ACTION act_Oper:
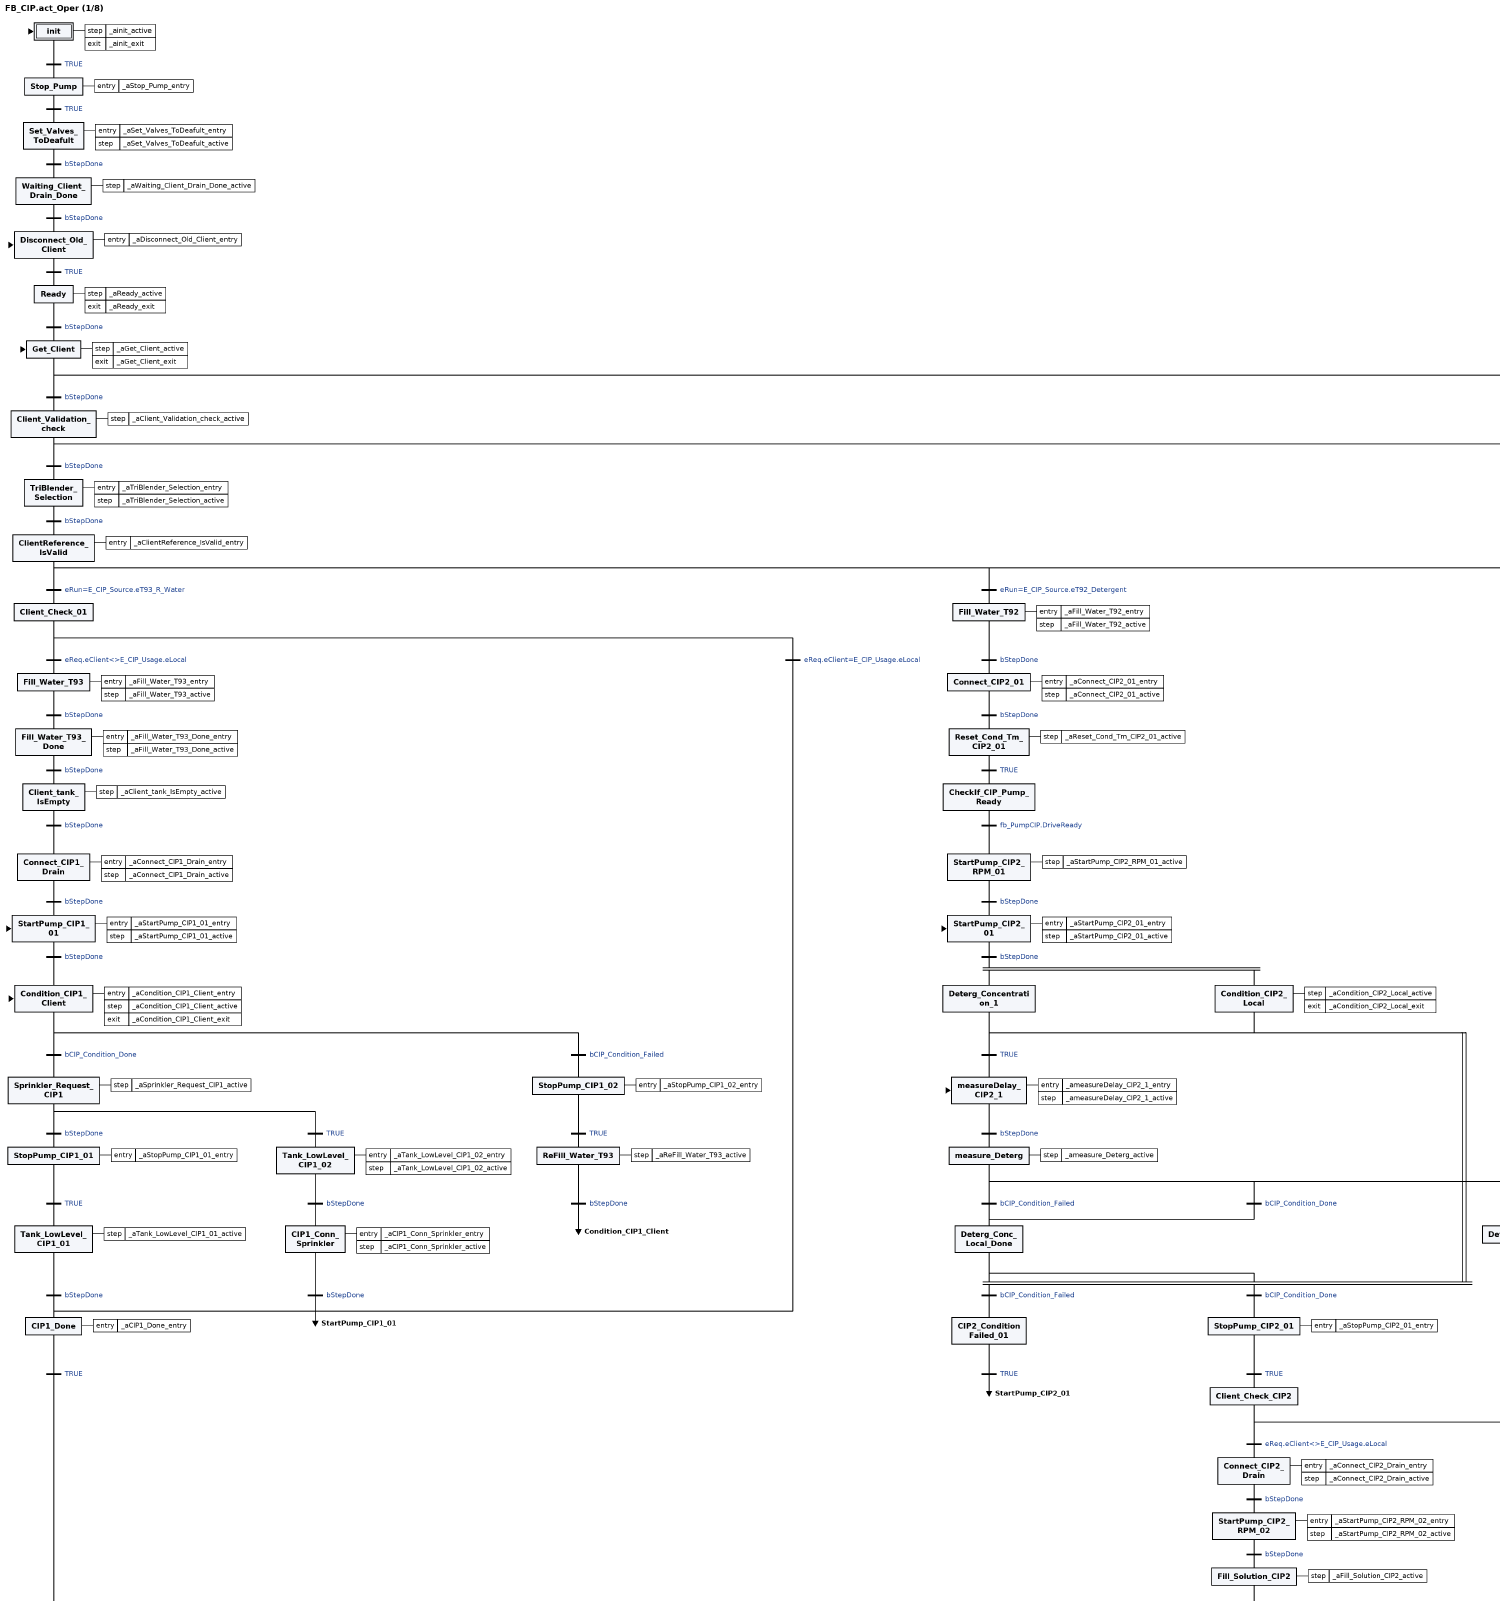
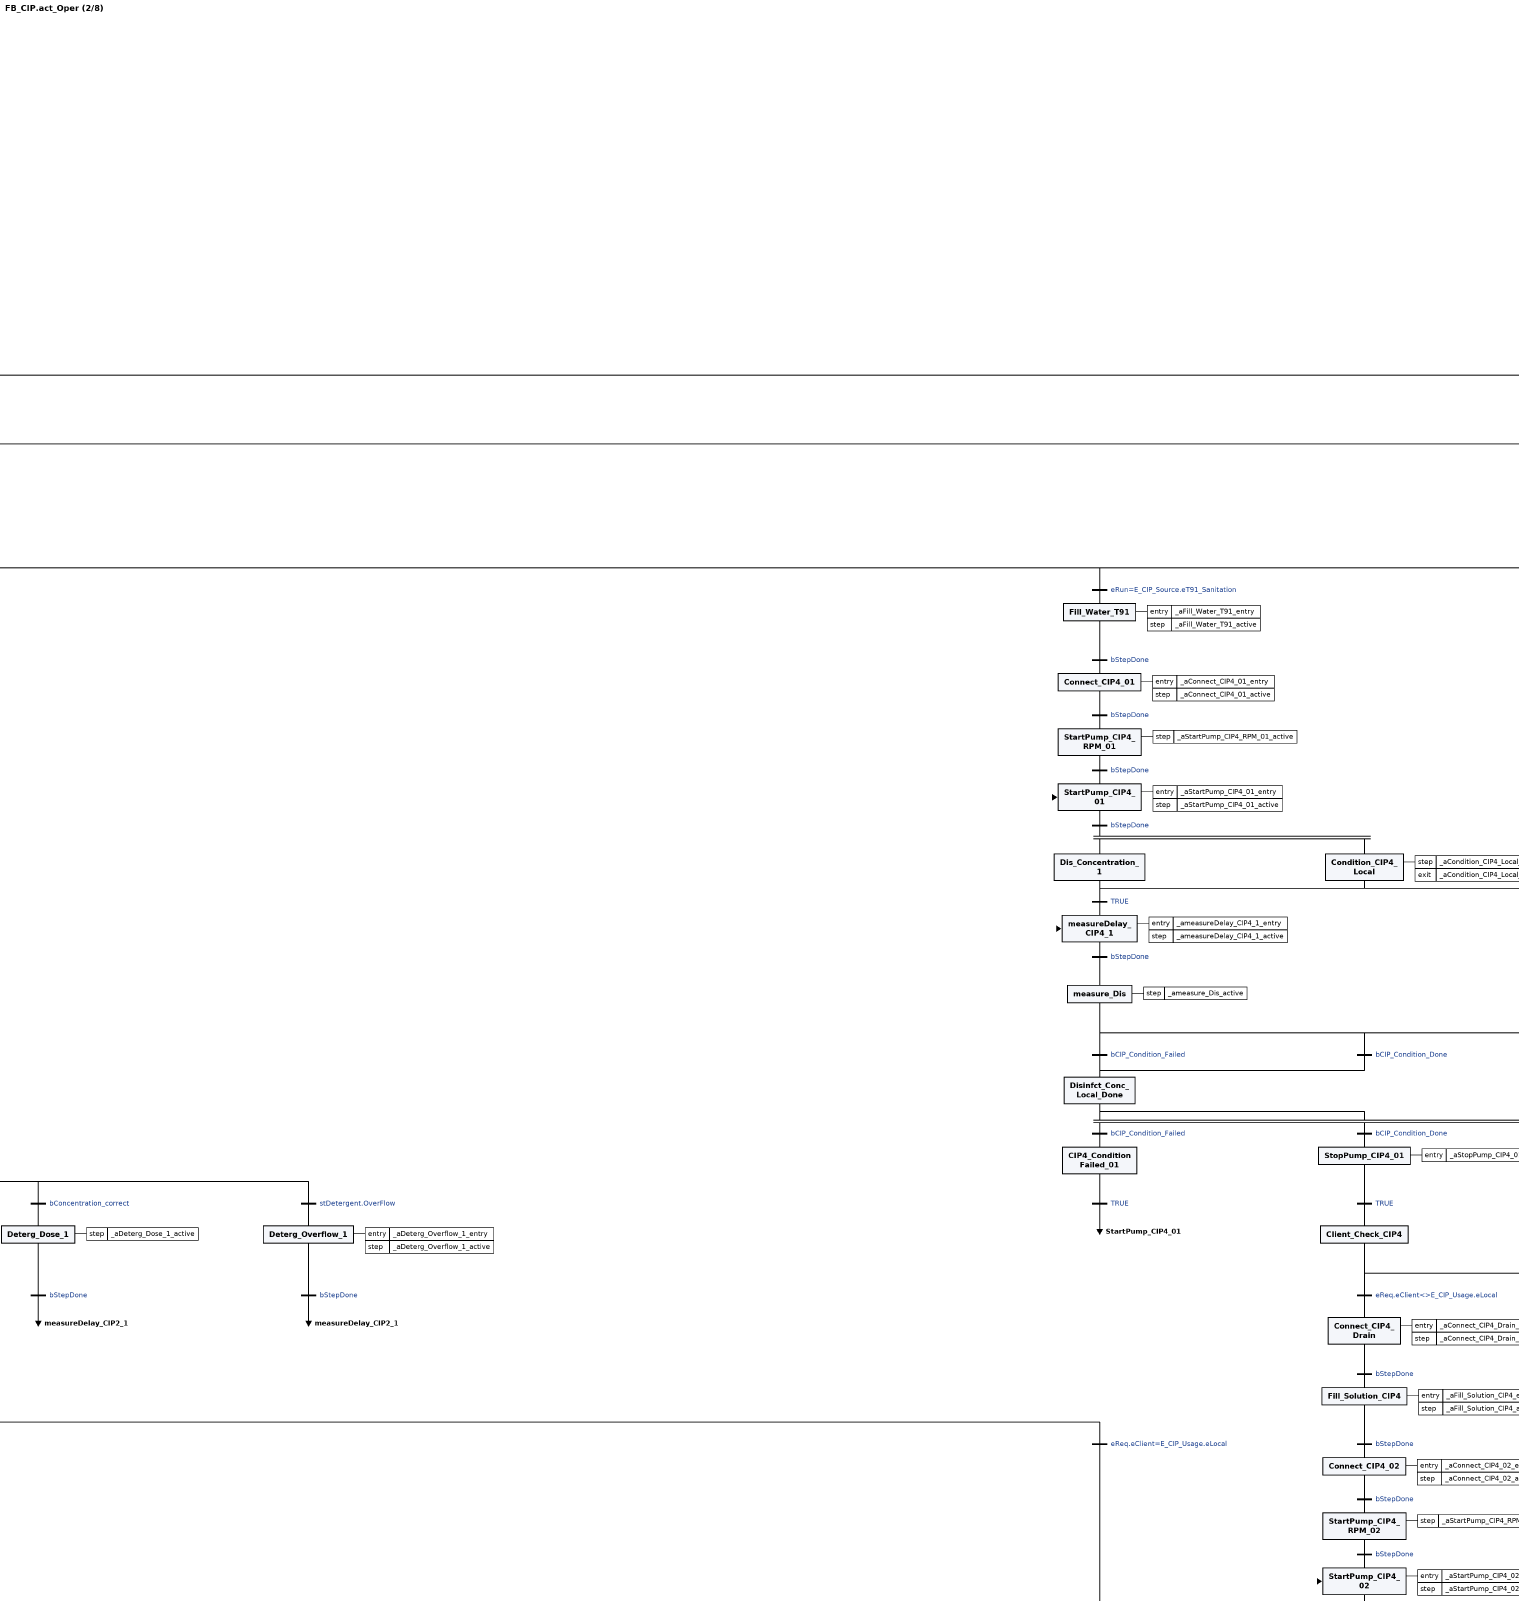
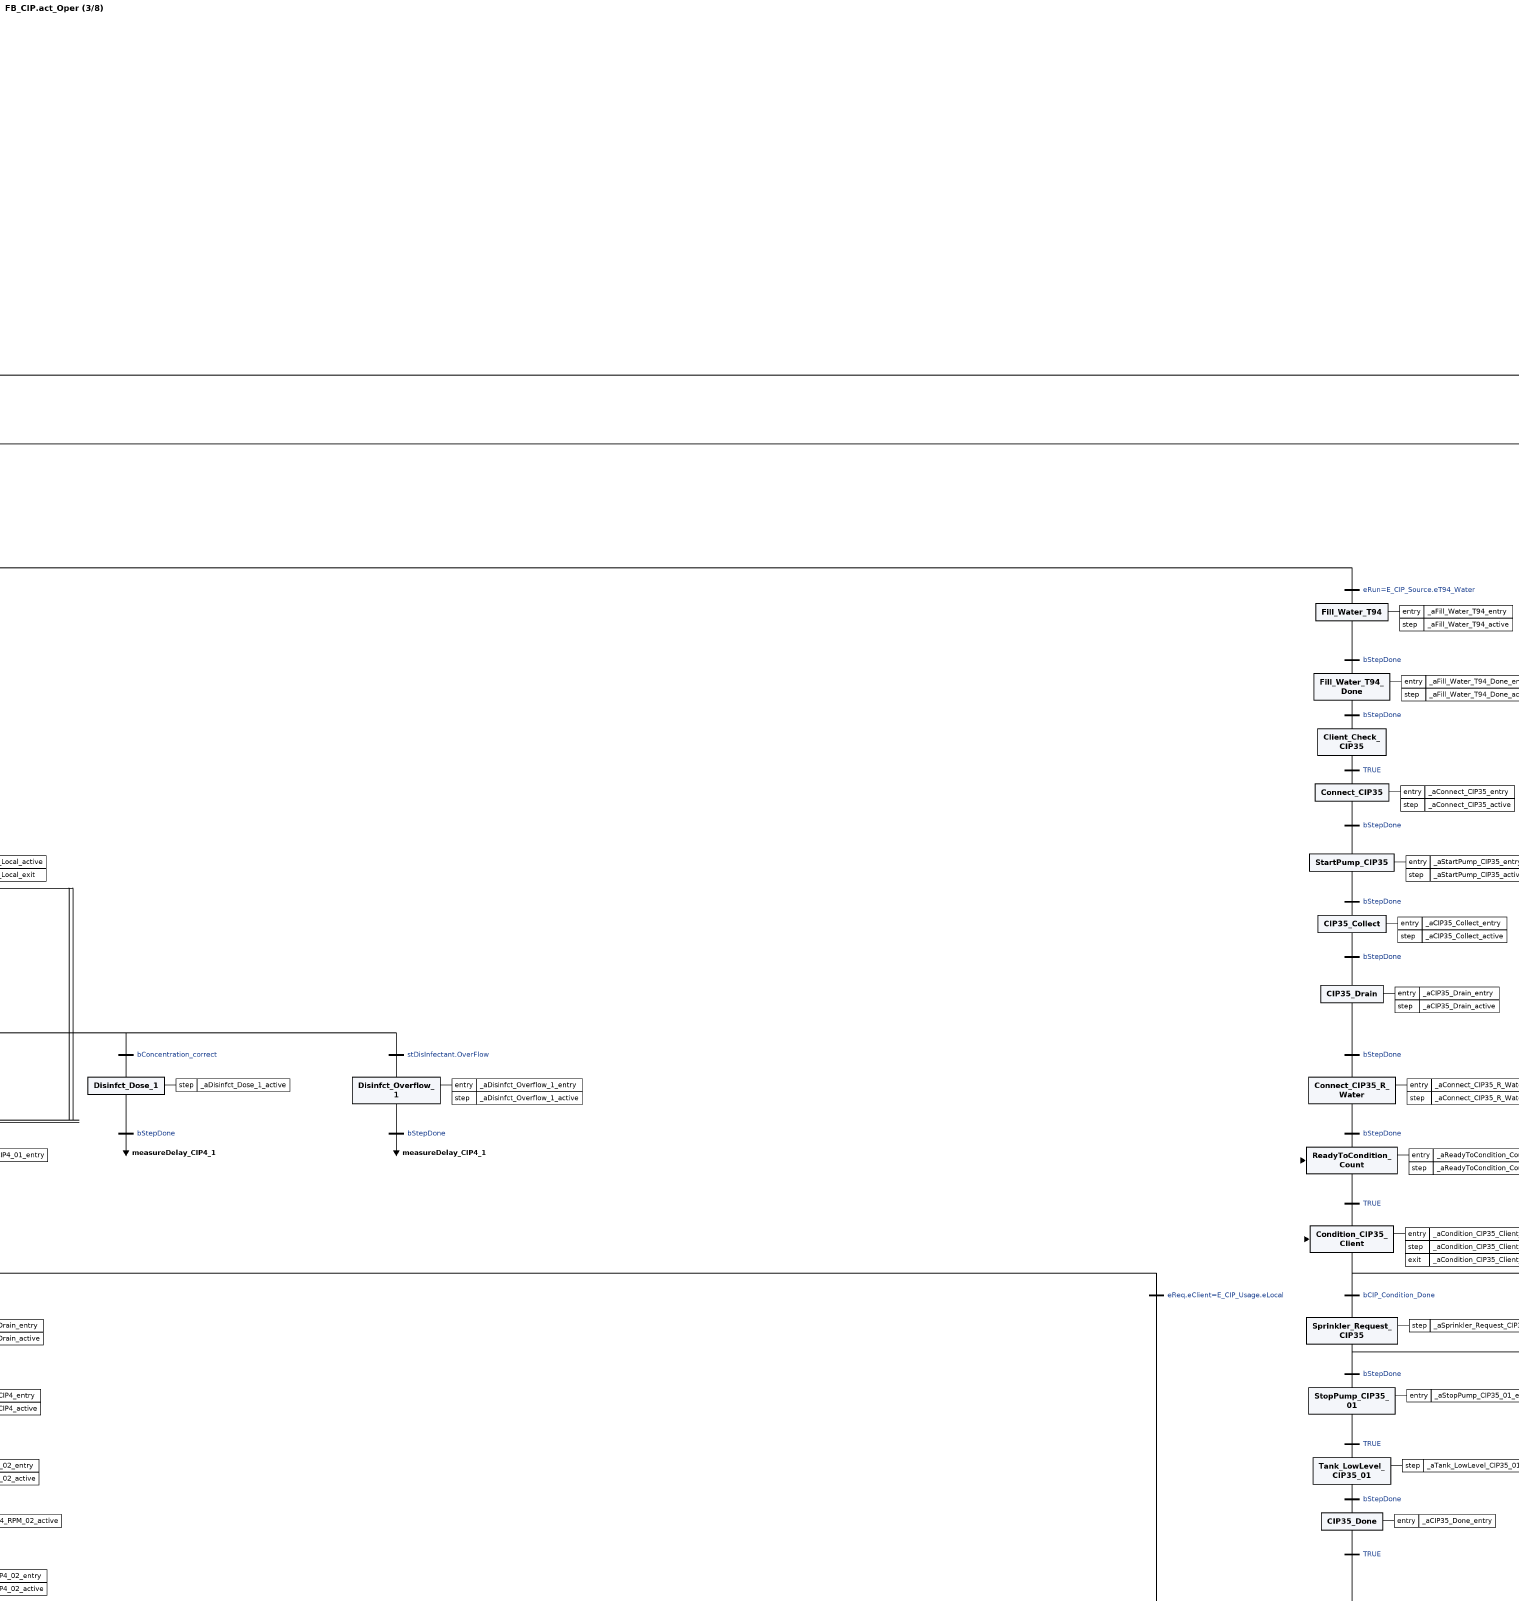
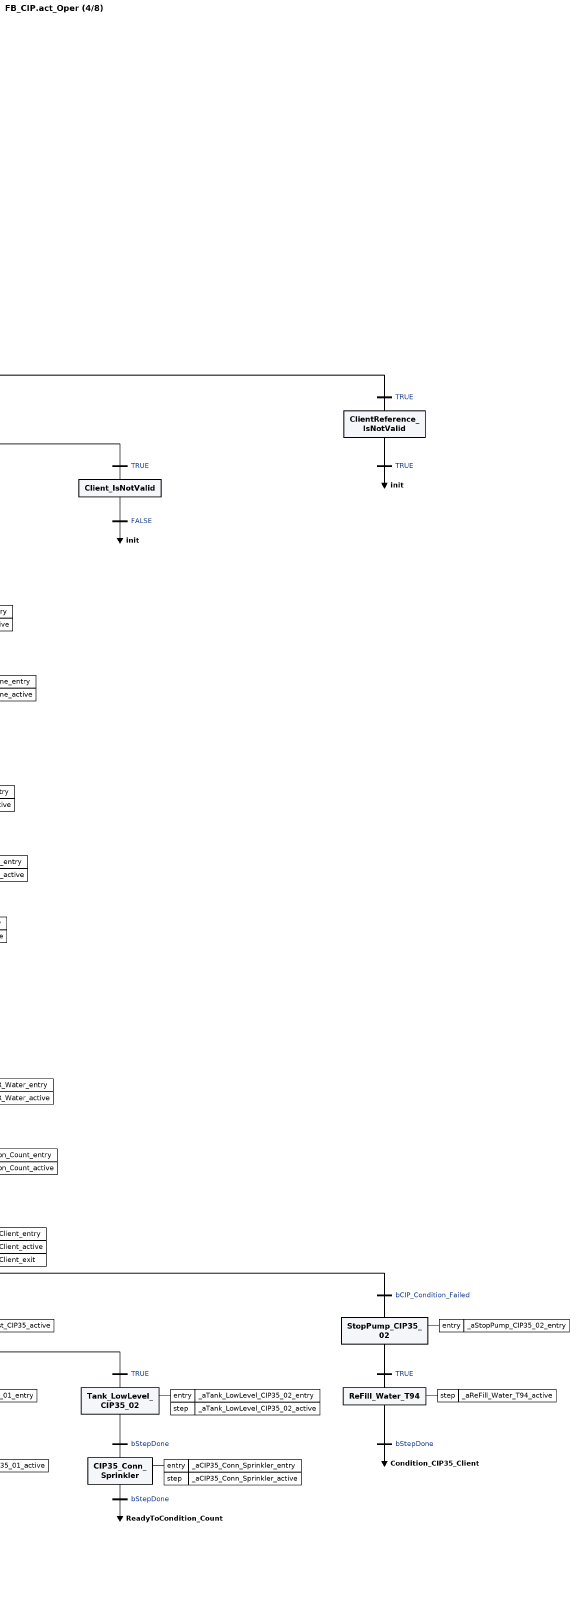
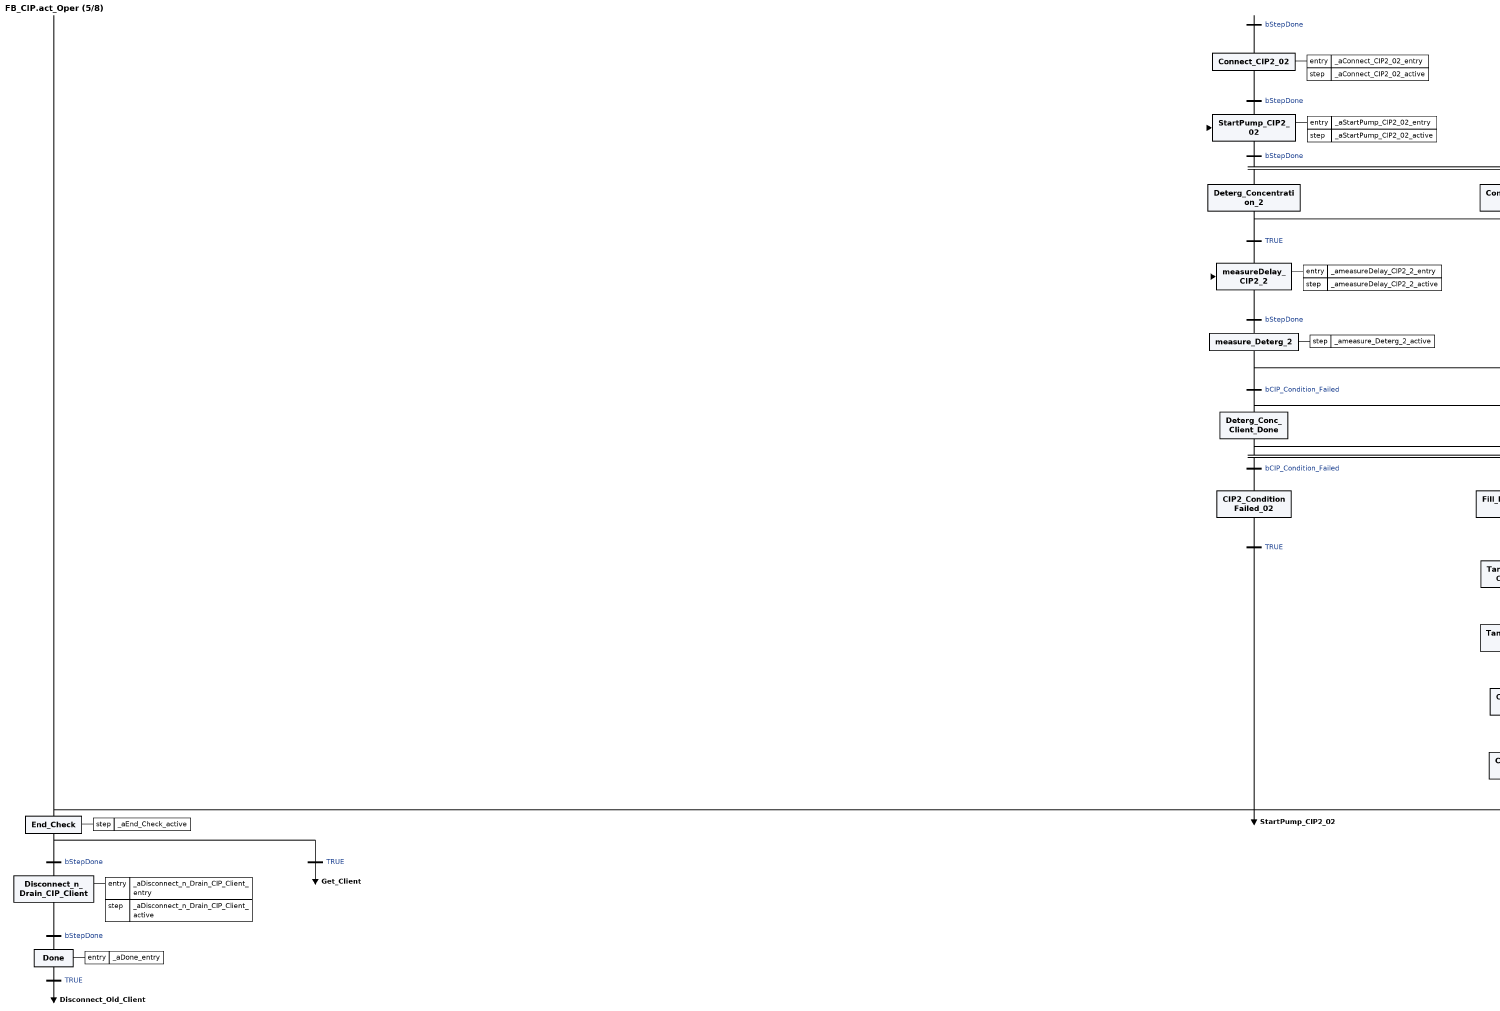
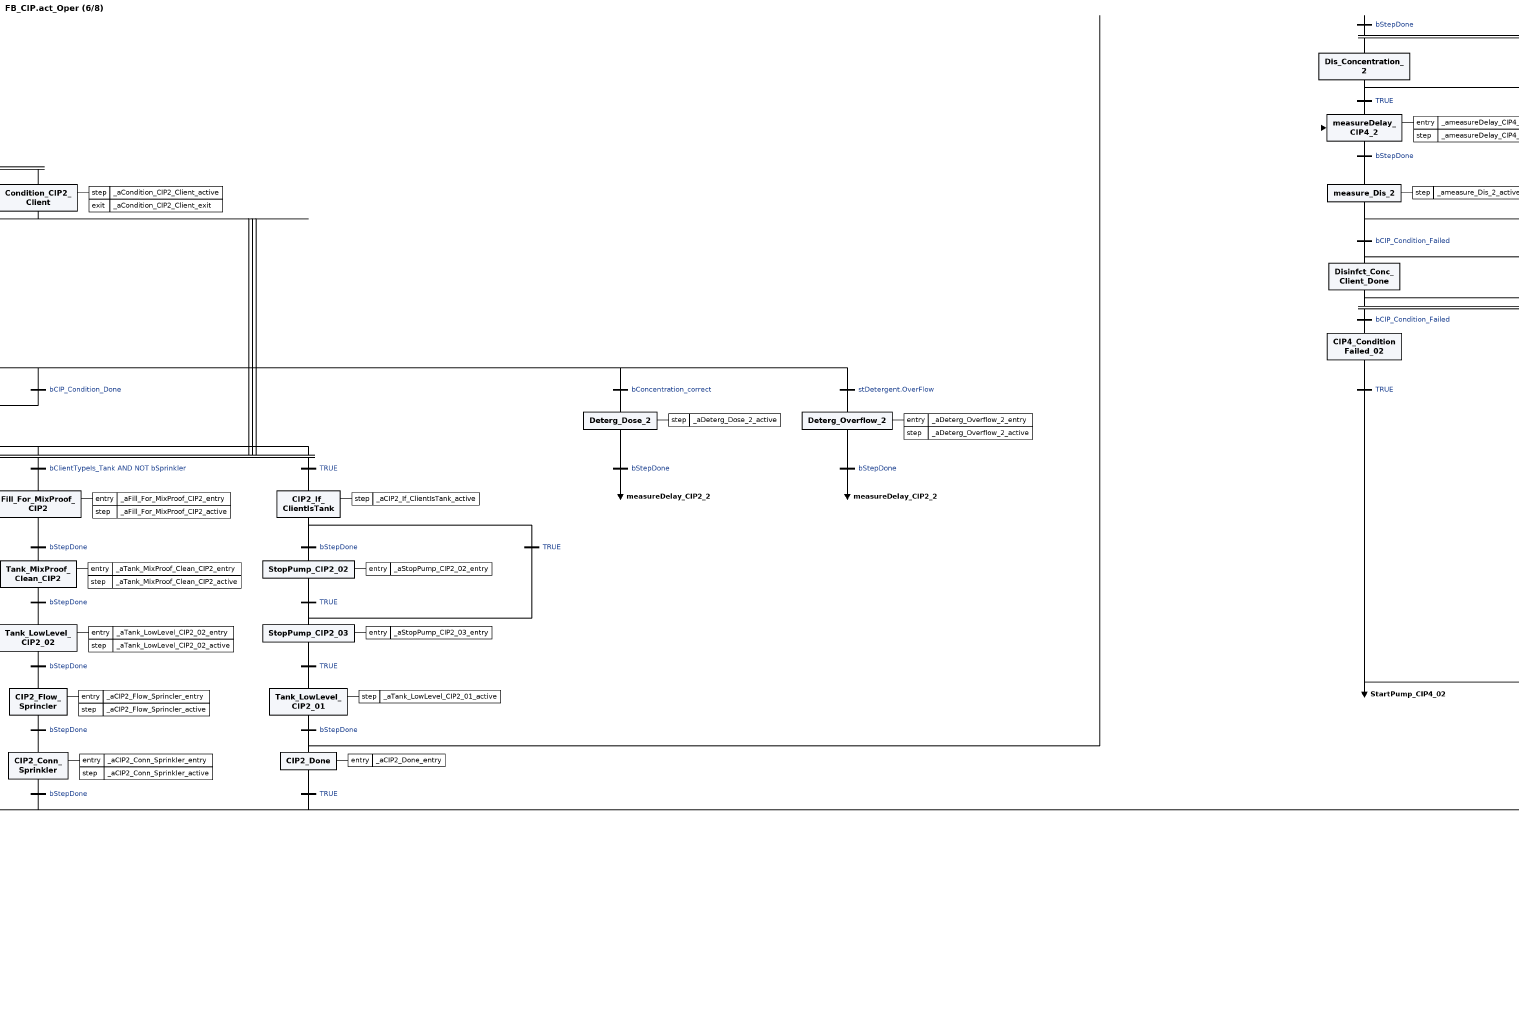
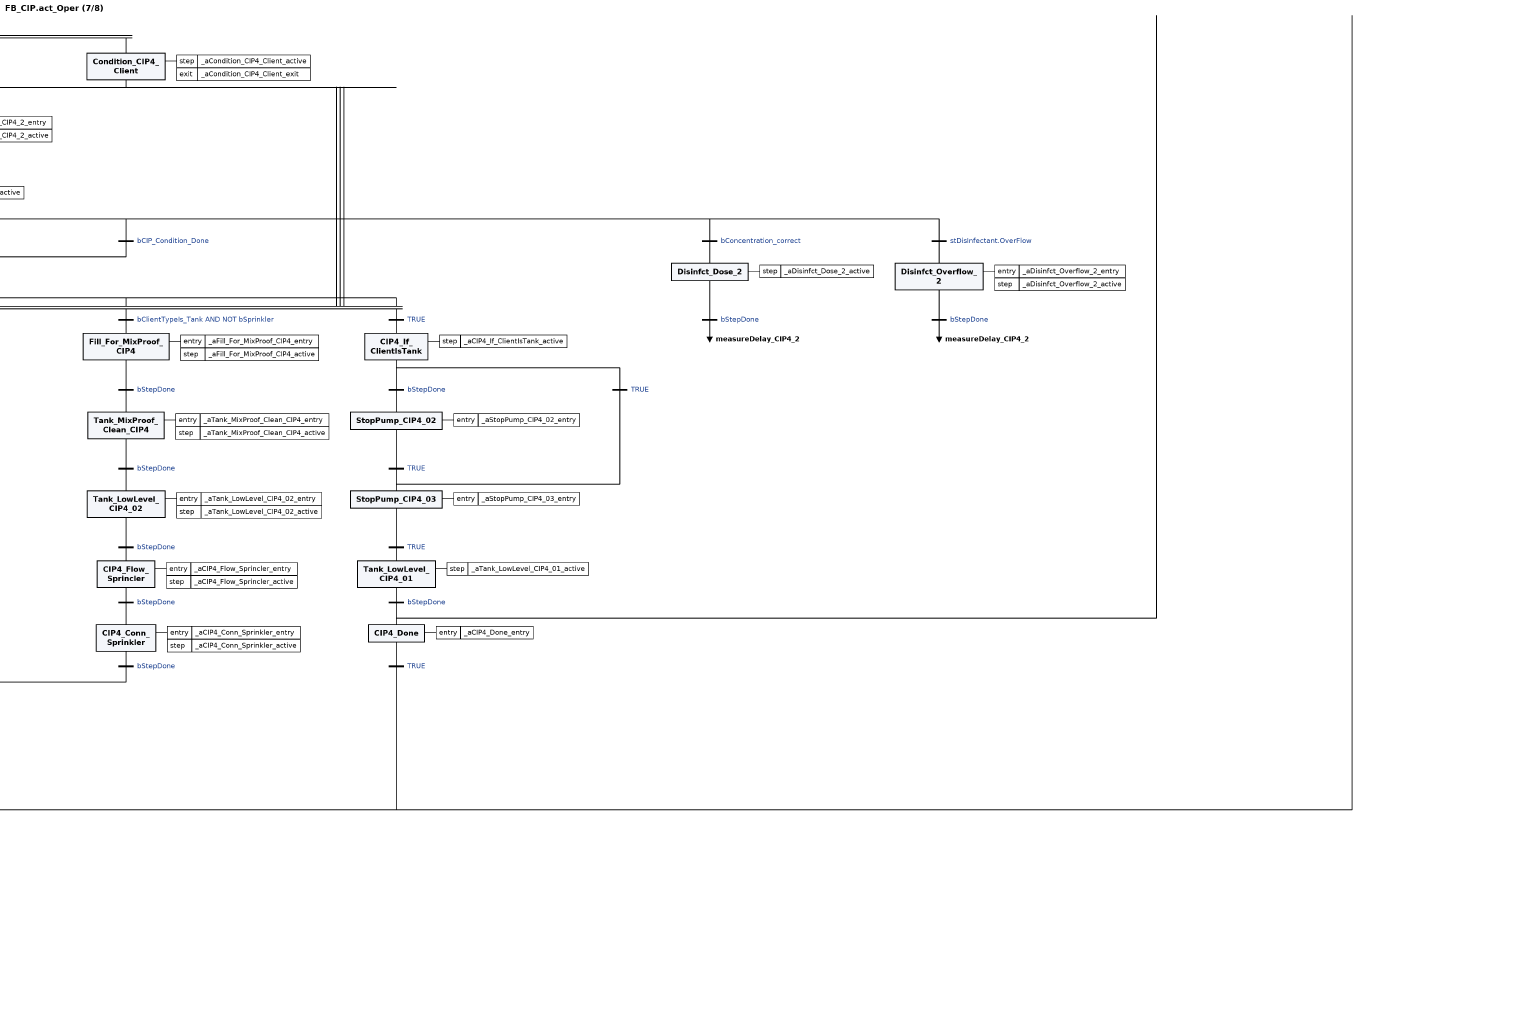
INITIAL_STEP init:
    _ainit_active(N);  // step action
    _ainit_exit(P0);  // exit action
END_STEP
TRANSITION FROM init TO Stop_Pump
    := TRUE;
END_TRANSITION
STEP Stop_Pump:
    _aStop_Pump_entry(P1);  // entry action
END_STEP
TRANSITION FROM Stop_Pump TO Set_Valves_ToDeafult
    := TRUE;
END_TRANSITION
STEP Set_Valves_ToDeafult:  // min time T#0.1s
    _aSet_Valves_ToDeafult_entry(P1);  // entry action
    _aSet_Valves_ToDeafult_active(N);  // step action
END_STEP
TRANSITION FROM Set_Valves_ToDeafult TO Waiting_Client_Drain_Done
    := bStepDone;
END_TRANSITION
STEP Waiting_Client_Drain_Done:  // min time T#0.1s
    _aWaiting_Client_Drain_Done_active(N);  // step action
END_STEP
TRANSITION FROM Waiting_Client_Drain_Done TO Disconnect_Old_Client
    := bStepDone;
END_TRANSITION
STEP Disconnect_Old_Client:
    _aDisconnect_Old_Client_entry(P1);  // entry action
END_STEP
TRANSITION FROM Disconnect_Old_Client TO Ready
    := TRUE;
END_TRANSITION
STEP Ready:
    _aReady_active(N);  // step action
    _aReady_exit(P0);  // exit action
END_STEP
TRANSITION FROM Ready TO Get_Client
    := bStepDone;
END_TRANSITION
STEP Get_Client:  // max time T#0.1s
    _aGet_Client_active(N);  // step action
    _aGet_Client_exit(P0);  // exit action
END_STEP
TRANSITION FROM Get_Client TO Client_Validation_check
    := bStepDone;
END_TRANSITION
TRANSITION FROM Get_Client TO ClientReference_IsNotValid
    := TRUE;
END_TRANSITION
STEP ClientReference_IsNotValid:  // min time T#2s
END_STEP
TRANSITION FROM ClientReference_IsNotValid TO init
    := TRUE;
END_TRANSITION
STEP Client_Validation_check:
    _aClient_Validation_check_active(N);  // step action
END_STEP
TRANSITION FROM Client_Validation_check TO TriBlender_Selection
    := bStepDone;
END_TRANSITION
STEP TriBlender_Selection:
    _aTriBlender_Selection_entry(P1);  // entry action
    _aTriBlender_Selection_active(N);  // step action
END_STEP
TRANSITION FROM TriBlender_Selection TO ClientReference_IsValid
    := bStepDone;
END_TRANSITION
TRANSITION FROM Client_Validation_check TO Client_IsNotValid
    := TRUE;
END_TRANSITION
STEP Client_IsNotValid:  // min time T#2s
END_STEP
TRANSITION FROM Client_IsNotValid TO init
    := FALSE;
END_TRANSITION
STEP ClientReference_IsValid:
    _aClientReference_IsValid_entry(P1);  // entry action
END_STEP
TRANSITION FROM ClientReference_IsValid TO Client_Check_01
    := eRun=E_CIP_Source.eT93_R_Water;
END_TRANSITION
// macro R_Water begins
STEP Client_Check_01:
END_STEP
TRANSITION FROM Client_Check_01 TO Fill_Water_T93
    := eReq.eClient<>E_CIP_Usage.eLocal;
END_TRANSITION
STEP Fill_Water_T93:
    _aFill_Water_T93_entry(P1);  // entry action
    _aFill_Water_T93_active(N);  // step action
END_STEP
TRANSITION FROM Fill_Water_T93 TO Fill_Water_T93_Done
    := bStepDone;
END_TRANSITION
STEP Fill_Water_T93_Done:
    _aFill_Water_T93_Done_entry(P1);  // entry action
    _aFill_Water_T93_Done_active(N);  // step action
END_STEP
TRANSITION FROM Fill_Water_T93_Done TO Client_tank_IsEmpty
    := bStepDone;
END_TRANSITION
STEP Client_tank_IsEmpty:  // min time T#5s
    _aClient_tank_IsEmpty_active(N);  // step action
END_STEP
TRANSITION FROM Client_tank_IsEmpty TO Connect_CIP1_Drain
    := bStepDone;
END_TRANSITION
STEP Connect_CIP1_Drain:
    _aConnect_CIP1_Drain_entry(P1);  // entry action
    _aConnect_CIP1_Drain_active(N);  // step action
END_STEP
TRANSITION FROM Connect_CIP1_Drain TO StartPump_CIP1_01
    := bStepDone;
END_TRANSITION
STEP StartPump_CIP1_01:
    _aStartPump_CIP1_01_entry(P1);  // entry action
    _aStartPump_CIP1_01_active(N);  // step action
END_STEP
TRANSITION FROM StartPump_CIP1_01 TO Condition_CIP1_Client
    := bStepDone;
END_TRANSITION
STEP Condition_CIP1_Client:
    _aCondition_CIP1_Client_entry(P1);  // entry action
    _aCondition_CIP1_Client_active(N);  // step action
    _aCondition_CIP1_Client_exit(P0);  // exit action
END_STEP
TRANSITION FROM Condition_CIP1_Client TO Sprinkler_Request_CIP1
    := bCIP_Condition_Done;
END_TRANSITION
STEP Sprinkler_Request_CIP1:
    _aSprinkler_Request_CIP1_active(N);  // step action
END_STEP
TRANSITION FROM Sprinkler_Request_CIP1 TO StopPump_CIP1_01
    := bStepDone;
END_TRANSITION
STEP StopPump_CIP1_01:
    _aStopPump_CIP1_01_entry(P1);  // entry action
END_STEP
TRANSITION FROM StopPump_CIP1_01 TO Tank_LowLevel_CIP1_01
    := TRUE;
END_TRANSITION
STEP Tank_LowLevel_CIP1_01:
    _aTank_LowLevel_CIP1_01_active(N);  // step action
END_STEP
TRANSITION FROM Tank_LowLevel_CIP1_01 TO CIP1_Done
    := bStepDone;
END_TRANSITION
TRANSITION FROM Sprinkler_Request_CIP1 TO Tank_LowLevel_CIP1_02
    := TRUE;
END_TRANSITION
STEP Tank_LowLevel_CIP1_02:
    _aTank_LowLevel_CIP1_02_entry(P1);  // entry action
    _aTank_LowLevel_CIP1_02_active(N);  // step action
END_STEP
TRANSITION FROM Tank_LowLevel_CIP1_02 TO CIP1_Conn_Sprinkler
    := bStepDone;
END_TRANSITION
STEP CIP1_Conn_Sprinkler:
    _aCIP1_Conn_Sprinkler_entry(P1);  // entry action
    _aCIP1_Conn_Sprinkler_active(N);  // step action
END_STEP
TRANSITION FROM CIP1_Conn_Sprinkler TO StartPump_CIP1_01
    := bStepDone;
END_TRANSITION
TRANSITION FROM Condition_CIP1_Client TO StopPump_CIP1_02
    := bCIP_Condition_Failed;
END_TRANSITION
STEP StopPump_CIP1_02:
    _aStopPump_CIP1_02_entry(P1);  // entry action
END_STEP
TRANSITION FROM StopPump_CIP1_02 TO ReFill_Water_T93
    := TRUE;
END_TRANSITION
STEP ReFill_Water_T93:
    _aReFill_Water_T93_active(N);  // step action
END_STEP
TRANSITION FROM ReFill_Water_T93 TO Condition_CIP1_Client
    := bStepDone;
END_TRANSITION
TRANSITION FROM Client_Check_01 TO CIP1_Done
    := eReq.eClient=E_CIP_Usage.eLocal;
END_TRANSITION
STEP CIP1_Done:  // min time T#2s
    _aCIP1_Done_entry(P1);  // entry action
END_STEP
TRANSITION FROM CIP1_Done TO End_Check
    := TRUE;
END_TRANSITION
TRANSITION FROM ClientReference_IsValid TO Fill_Water_T92
    := eRun=E_CIP_Source.eT92_Detergent;
END_TRANSITION
// macro Detergent begins
STEP Fill_Water_T92:
    _aFill_Water_T92_entry(P1);  // entry action
    _aFill_Water_T92_active(N);  // step action
END_STEP
TRANSITION FROM Fill_Water_T92 TO Connect_CIP2_01
    := bStepDone;
END_TRANSITION
STEP Connect_CIP2_01:
    _aConnect_CIP2_01_entry(P1);  // entry action
    _aConnect_CIP2_01_active(N);  // step action
END_STEP
TRANSITION FROM Connect_CIP2_01 TO Reset_Cond_Tm_CIP2_01
    := bStepDone;
END_TRANSITION
STEP Reset_Cond_Tm_CIP2_01:
    _aReset_Cond_Tm_CIP2_01_active(N);  // step action
END_STEP
TRANSITION FROM Reset_Cond_Tm_CIP2_01 TO CheckIf_CIP_Pump_Ready
    := TRUE;
END_TRANSITION
STEP CheckIf_CIP_Pump_Ready:
END_STEP
TRANSITION FROM CheckIf_CIP_Pump_Ready TO StartPump_CIP2_RPM_01
    := fb_PumpCIP.DriveReady;
END_TRANSITION
STEP StartPump_CIP2_RPM_01:
    _aStartPump_CIP2_RPM_01_active(N);  // step action
END_STEP
TRANSITION FROM StartPump_CIP2_RPM_01 TO StartPump_CIP2_01
    := bStepDone;
END_TRANSITION
STEP StartPump_CIP2_01:  // min time T#2s
    _aStartPump_CIP2_01_entry(P1);  // entry action
    _aStartPump_CIP2_01_active(N);  // step action
END_STEP
TRANSITION FROM StartPump_CIP2_01 TO (Deterg_Concentration_1, Condition_CIP2_Local)
    := bStepDone;
END_TRANSITION
STEP Deterg_Concentration_1:
END_STEP
TRANSITION FROM Deterg_Concentration_1 TO measureDelay_CIP2_1
    := TRUE;
END_TRANSITION
STEP measureDelay_CIP2_1:
    _ameasureDelay_CIP2_1_entry(P1);  // entry action
    _ameasureDelay_CIP2_1_active(N);  // step action
END_STEP
TRANSITION FROM measureDelay_CIP2_1 TO measure_Deterg
    := bStepDone;
END_TRANSITION
STEP measure_Deterg:  // min time t#1s
    _ameasure_Deterg_active(N);  // step action
END_STEP
TRANSITION FROM measure_Deterg TO Deterg_Conc_Local_Done
    := bCIP_Condition_Failed;
END_TRANSITION
TRANSITION FROM measure_Deterg TO Deterg_Conc_Local_Done
    := bCIP_Condition_Done;
END_TRANSITION
TRANSITION FROM measure_Deterg TO Deterg_Dose_1
    := bConcentration_correct;
END_TRANSITION
STEP Deterg_Dose_1:
    _aDeterg_Dose_1_active(N);  // step action
END_STEP
TRANSITION FROM Deterg_Dose_1 TO measureDelay_CIP2_1
    := bStepDone;
END_TRANSITION
TRANSITION FROM measure_Deterg TO Deterg_Overflow_1
    := stDetergent.OverFlow;
END_TRANSITION
STEP Deterg_Overflow_1:
    _aDeterg_Overflow_1_entry(P1);  // entry action
    _aDeterg_Overflow_1_active(N);  // step action
END_STEP
TRANSITION FROM Deterg_Overflow_1 TO measureDelay_CIP2_1
    := bStepDone;
END_TRANSITION
STEP Deterg_Conc_Local_Done:
END_STEP
STEP Condition_CIP2_Local:
    _aCondition_CIP2_Local_active(N);  // step action
    _aCondition_CIP2_Local_exit(P0);  // exit action
END_STEP
TRANSITION FROM (Deterg_Conc_Local_Done, Condition_CIP2_Local) TO CIP2_ConditionFailed_01
    := bCIP_Condition_Failed;
END_TRANSITION
STEP CIP2_ConditionFailed_01:
END_STEP
TRANSITION FROM CIP2_ConditionFailed_01 TO StartPump_CIP2_01
    := TRUE;
END_TRANSITION
TRANSITION FROM (Deterg_Conc_Local_Done, Condition_CIP2_Local) TO StopPump_CIP2_01
    := bCIP_Condition_Done;
END_TRANSITION
STEP StopPump_CIP2_01:
    _aStopPump_CIP2_01_entry(P1);  // entry action
END_STEP
TRANSITION FROM StopPump_CIP2_01 TO Client_Check_CIP2
    := TRUE;
END_TRANSITION
STEP Client_Check_CIP2:
END_STEP
TRANSITION FROM Client_Check_CIP2 TO Connect_CIP2_Drain
    := eReq.eClient<>E_CIP_Usage.eLocal;
END_TRANSITION
STEP Connect_CIP2_Drain:
    _aConnect_CIP2_Drain_entry(P1);  // entry action
    _aConnect_CIP2_Drain_active(N);  // step action
END_STEP
TRANSITION FROM Connect_CIP2_Drain TO StartPump_CIP2_RPM_02
    := bStepDone;
END_TRANSITION
STEP StartPump_CIP2_RPM_02:
    _aStartPump_CIP2_RPM_02_entry(P1);  // entry action
    _aStartPump_CIP2_RPM_02_active(N);  // step action
END_STEP
TRANSITION FROM StartPump_CIP2_RPM_02 TO Fill_Solution_CIP2
    := bStepDone;
END_TRANSITION
STEP Fill_Solution_CIP2:
    _aFill_Solution_CIP2_active(N);  // step action
END_STEP
TRANSITION FROM Fill_Solution_CIP2 TO Connect_CIP2_02
    := bStepDone;
END_TRANSITION
STEP Connect_CIP2_02:
    _aConnect_CIP2_02_entry(P1);  // entry action
    _aConnect_CIP2_02_active(N);  // step action
END_STEP
TRANSITION FROM Connect_CIP2_02 TO StartPump_CIP2_02
    := bStepDone;
END_TRANSITION
STEP StartPump_CIP2_02:  // min time T#2s
    _aStartPump_CIP2_02_entry(P1);  // entry action
    _aStartPump_CIP2_02_active(N);  // step action
END_STEP
TRANSITION FROM StartPump_CIP2_02 TO (Deterg_Concentration_2, Condition_CIP2_Client)
    := bStepDone;
END_TRANSITION
STEP Deterg_Concentration_2:
END_STEP
TRANSITION FROM Deterg_Concentration_2 TO measureDelay_CIP2_2
    := TRUE;
END_TRANSITION
STEP measureDelay_CIP2_2:
    _ameasureDelay_CIP2_2_entry(P1);  // entry action
    _ameasureDelay_CIP2_2_active(N);  // step action
END_STEP
TRANSITION FROM measureDelay_CIP2_2 TO measure_Deterg_2
    := bStepDone;
END_TRANSITION
STEP measure_Deterg_2:  // min time t#1s
    _ameasure_Deterg_2_active(N);  // step action
END_STEP
TRANSITION FROM measure_Deterg_2 TO Deterg_Conc_Client_Done
    := bCIP_Condition_Failed;
END_TRANSITION
TRANSITION FROM measure_Deterg_2 TO Deterg_Conc_Client_Done
    := bCIP_Condition_Done;
END_TRANSITION
TRANSITION FROM measure_Deterg_2 TO Deterg_Dose_2
    := bConcentration_correct;
END_TRANSITION
STEP Deterg_Dose_2:
    _aDeterg_Dose_2_active(N);  // step action
END_STEP
TRANSITION FROM Deterg_Dose_2 TO measureDelay_CIP2_2
    := bStepDone;
END_TRANSITION
TRANSITION FROM measure_Deterg_2 TO Deterg_Overflow_2
    := stDetergent.OverFlow;
END_TRANSITION
STEP Deterg_Overflow_2:
    _aDeterg_Overflow_2_entry(P1);  // entry action
    _aDeterg_Overflow_2_active(N);  // step action
END_STEP
TRANSITION FROM Deterg_Overflow_2 TO measureDelay_CIP2_2
    := bStepDone;
END_TRANSITION
STEP Deterg_Conc_Client_Done:
END_STEP
STEP Condition_CIP2_Client:
    _aCondition_CIP2_Client_active(N);  // step action
    _aCondition_CIP2_Client_exit(P0);  // exit action
END_STEP
TRANSITION FROM (Deterg_Conc_Client_Done, Condition_CIP2_Client) TO CIP2_ConditionFailed_02
    := bCIP_Condition_Failed;
END_TRANSITION
STEP CIP2_ConditionFailed_02:
END_STEP
TRANSITION FROM CIP2_ConditionFailed_02 TO StartPump_CIP2_02
    := TRUE;
END_TRANSITION
TRANSITION FROM (Deterg_Conc_Client_Done, Condition_CIP2_Client) TO Fill_For_MixProof_CIP2
    := bClientTypeIs_Tank AND NOT bSprinkler;
END_TRANSITION
STEP Fill_For_MixProof_CIP2:
    _aFill_For_MixProof_CIP2_entry(P1);  // entry action
    _aFill_For_MixProof_CIP2_active(N);  // step action
END_STEP
TRANSITION FROM Fill_For_MixProof_CIP2 TO Tank_MixProof_Clean_CIP2
    := bStepDone;
END_TRANSITION
STEP Tank_MixProof_Clean_CIP2:
    _aTank_MixProof_Clean_CIP2_entry(P1);  // entry action
    _aTank_MixProof_Clean_CIP2_active(N);  // step action
END_STEP
TRANSITION FROM Tank_MixProof_Clean_CIP2 TO Tank_LowLevel_CIP2_02
    := bStepDone;
END_TRANSITION
STEP Tank_LowLevel_CIP2_02:
    _aTank_LowLevel_CIP2_02_entry(P1);  // entry action
    _aTank_LowLevel_CIP2_02_active(N);  // step action
END_STEP
TRANSITION FROM Tank_LowLevel_CIP2_02 TO CIP2_Flow_Sprincler
    := bStepDone;
END_TRANSITION
STEP CIP2_Flow_Sprincler:
    _aCIP2_Flow_Sprincler_entry(P1);  // entry action
    _aCIP2_Flow_Sprincler_active(N);  // step action
END_STEP
TRANSITION FROM CIP2_Flow_Sprincler TO CIP2_Conn_Sprinkler
    := bStepDone;
END_TRANSITION
STEP CIP2_Conn_Sprinkler:
    _aCIP2_Conn_Sprinkler_entry(P1);  // entry action
    _aCIP2_Conn_Sprinkler_active(N);  // step action
END_STEP
TRANSITION FROM CIP2_Conn_Sprinkler TO StartPump_CIP2_02
    := bStepDone;
END_TRANSITION
TRANSITION FROM (Deterg_Conc_Client_Done, Condition_CIP2_Client) TO CIP2_If_ClientIsTank
    := TRUE;
END_TRANSITION
STEP CIP2_If_ClientIsTank:
    _aCIP2_If_ClientIsTank_active(N);  // step action
END_STEP
TRANSITION FROM CIP2_If_ClientIsTank TO StopPump_CIP2_02
    := bStepDone;
END_TRANSITION
STEP StopPump_CIP2_02:
    _aStopPump_CIP2_02_entry(P1);  // entry action
END_STEP
TRANSITION FROM StopPump_CIP2_02 TO StopPump_CIP2_03
    := TRUE;
END_TRANSITION
TRANSITION FROM CIP2_If_ClientIsTank TO StopPump_CIP2_03
    := TRUE;
END_TRANSITION
STEP StopPump_CIP2_03:
    _aStopPump_CIP2_03_entry(P1);  // entry action
END_STEP
TRANSITION FROM StopPump_CIP2_03 TO Tank_LowLevel_CIP2_01
    := TRUE;
END_TRANSITION
STEP Tank_LowLevel_CIP2_01:
    _aTank_LowLevel_CIP2_01_active(N);  // step action
END_STEP
TRANSITION FROM Tank_LowLevel_CIP2_01 TO CIP2_Done
    := bStepDone;
END_TRANSITION
TRANSITION FROM Client_Check_CIP2 TO CIP2_Done
    := eReq.eClient=E_CIP_Usage.eLocal;
END_TRANSITION
STEP CIP2_Done:  // min time T#2s
    _aCIP2_Done_entry(P1);  // entry action
END_STEP
TRANSITION FROM CIP2_Done TO End_Check
    := TRUE;
END_TRANSITION
TRANSITION FROM ClientReference_IsValid TO Fill_Water_T91
    := eRun=E_CIP_Source.eT91_Sanitation;
END_TRANSITION
// macro DisInfection begins
STEP Fill_Water_T91:
    _aFill_Water_T91_entry(P1);  // entry action
    _aFill_Water_T91_active(N);  // step action
END_STEP
TRANSITION FROM Fill_Water_T91 TO Connect_CIP4_01
    := bStepDone;
END_TRANSITION
STEP Connect_CIP4_01:
    _aConnect_CIP4_01_entry(P1);  // entry action
    _aConnect_CIP4_01_active(N);  // step action
END_STEP
TRANSITION FROM Connect_CIP4_01 TO StartPump_CIP4_RPM_01
    := bStepDone;
END_TRANSITION
STEP StartPump_CIP4_RPM_01:
    _aStartPump_CIP4_RPM_01_active(N);  // step action
END_STEP
TRANSITION FROM StartPump_CIP4_RPM_01 TO StartPump_CIP4_01
    := bStepDone;
END_TRANSITION
STEP StartPump_CIP4_01:  // min time T#3s
    _aStartPump_CIP4_01_entry(P1);  // entry action
    _aStartPump_CIP4_01_active(N);  // step action
END_STEP
TRANSITION FROM StartPump_CIP4_01 TO (Dis_Concentration_1, Condition_CIP4_Local)
    := bStepDone;
END_TRANSITION
STEP Dis_Concentration_1:
END_STEP
TRANSITION FROM Dis_Concentration_1 TO measureDelay_CIP4_1
    := TRUE;
END_TRANSITION
STEP measureDelay_CIP4_1:
    _ameasureDelay_CIP4_1_entry(P1);  // entry action
    _ameasureDelay_CIP4_1_active(N);  // step action
END_STEP
TRANSITION FROM measureDelay_CIP4_1 TO measure_Dis
    := bStepDone;
END_TRANSITION
STEP measure_Dis:  // min time t#1s
    _ameasure_Dis_active(N);  // step action
END_STEP
TRANSITION FROM measure_Dis TO Disinfct_Conc_Local_Done
    := bCIP_Condition_Failed;
END_TRANSITION
TRANSITION FROM measure_Dis TO Disinfct_Conc_Local_Done
    := bCIP_Condition_Done;
END_TRANSITION
TRANSITION FROM measure_Dis TO Disinfct_Dose_1
    := bConcentration_correct;
END_TRANSITION
STEP Disinfct_Dose_1:
    _aDisinfct_Dose_1_active(N);  // step action
END_STEP
TRANSITION FROM Disinfct_Dose_1 TO measureDelay_CIP4_1
    := bStepDone;
END_TRANSITION
TRANSITION FROM measure_Dis TO Disinfct_Overflow_1
    := stDisInfectant.OverFlow;
END_TRANSITION
STEP Disinfct_Overflow_1:
    _aDisinfct_Overflow_1_entry(P1);  // entry action
    _aDisinfct_Overflow_1_active(N);  // step action
END_STEP
TRANSITION FROM Disinfct_Overflow_1 TO measureDelay_CIP4_1
    := bStepDone;
END_TRANSITION
STEP Disinfct_Conc_Local_Done:
END_STEP
STEP Condition_CIP4_Local:
    _aCondition_CIP4_Local_active(N);  // step action
    _aCondition_CIP4_Local_exit(P0);  // exit action
END_STEP
TRANSITION FROM (Disinfct_Conc_Local_Done, Condition_CIP4_Local) TO CIP4_ConditionFailed_01
    := bCIP_Condition_Failed;
END_TRANSITION
STEP CIP4_ConditionFailed_01:
END_STEP
TRANSITION FROM CIP4_ConditionFailed_01 TO StartPump_CIP4_01
    := TRUE;
END_TRANSITION
TRANSITION FROM (Disinfct_Conc_Local_Done, Condition_CIP4_Local) TO StopPump_CIP4_01
    := bCIP_Condition_Done;
END_TRANSITION
STEP StopPump_CIP4_01:  // min time T#5s
    _aStopPump_CIP4_01_entry(P1);  // entry action
END_STEP
TRANSITION FROM StopPump_CIP4_01 TO Client_Check_CIP4
    := TRUE;
END_TRANSITION
STEP Client_Check_CIP4:
END_STEP
TRANSITION FROM Client_Check_CIP4 TO Connect_CIP4_Drain
    := eReq.eClient<>E_CIP_Usage.eLocal;
END_TRANSITION
STEP Connect_CIP4_Drain:
    _aConnect_CIP4_Drain_entry(P1);  // entry action
    _aConnect_CIP4_Drain_active(N);  // step action
END_STEP
TRANSITION FROM Connect_CIP4_Drain TO Fill_Solution_CIP4
    := bStepDone;
END_TRANSITION
STEP Fill_Solution_CIP4:
    _aFill_Solution_CIP4_entry(P1);  // entry action
    _aFill_Solution_CIP4_active(N);  // step action
END_STEP
TRANSITION FROM Fill_Solution_CIP4 TO Connect_CIP4_02
    := bStepDone;
END_TRANSITION
STEP Connect_CIP4_02:
    _aConnect_CIP4_02_entry(P1);  // entry action
    _aConnect_CIP4_02_active(N);  // step action
END_STEP
TRANSITION FROM Connect_CIP4_02 TO StartPump_CIP4_RPM_02
    := bStepDone;
END_TRANSITION
STEP StartPump_CIP4_RPM_02:
    _aStartPump_CIP4_RPM_02_active(N);  // step action
END_STEP
TRANSITION FROM StartPump_CIP4_RPM_02 TO StartPump_CIP4_02
    := bStepDone;
END_TRANSITION
STEP StartPump_CIP4_02:  // min time T#1s
    _aStartPump_CIP4_02_entry(P1);  // entry action
    _aStartPump_CIP4_02_active(N);  // step action
END_STEP
TRANSITION FROM StartPump_CIP4_02 TO (Dis_Concentration_2, Condition_CIP4_Client)
    := bStepDone;
END_TRANSITION
STEP Dis_Concentration_2:
END_STEP
TRANSITION FROM Dis_Concentration_2 TO measureDelay_CIP4_2
    := TRUE;
END_TRANSITION
STEP measureDelay_CIP4_2:
    _ameasureDelay_CIP4_2_entry(P1);  // entry action
    _ameasureDelay_CIP4_2_active(N);  // step action
END_STEP
TRANSITION FROM measureDelay_CIP4_2 TO measure_Dis_2
    := bStepDone;
END_TRANSITION
STEP measure_Dis_2:  // min time t#1s
    _ameasure_Dis_2_active(N);  // step action
END_STEP
TRANSITION FROM measure_Dis_2 TO Disinfct_Conc_Client_Done
    := bCIP_Condition_Failed;
END_TRANSITION
TRANSITION FROM measure_Dis_2 TO Disinfct_Conc_Client_Done
    := bCIP_Condition_Done;
END_TRANSITION
TRANSITION FROM measure_Dis_2 TO Disinfct_Dose_2
    := bConcentration_correct;
END_TRANSITION
STEP Disinfct_Dose_2:
    _aDisinfct_Dose_2_active(N);  // step action
END_STEP
TRANSITION FROM Disinfct_Dose_2 TO measureDelay_CIP4_2
    := bStepDone;
END_TRANSITION
TRANSITION FROM measure_Dis_2 TO Disinfct_Overflow_2
    := stDisInfectant.OverFlow;
END_TRANSITION
STEP Disinfct_Overflow_2:
    _aDisinfct_Overflow_2_entry(P1);  // entry action
    _aDisinfct_Overflow_2_active(N);  // step action
END_STEP
TRANSITION FROM Disinfct_Overflow_2 TO measureDelay_CIP4_2
    := bStepDone;
END_TRANSITION
STEP Disinfct_Conc_Client_Done:
END_STEP
STEP Condition_CIP4_Client:
    _aCondition_CIP4_Client_active(N);  // step action
    _aCondition_CIP4_Client_exit(P0);  // exit action
END_STEP
TRANSITION FROM (Disinfct_Conc_Client_Done, Condition_CIP4_Client) TO CIP4_ConditionFailed_02
    := bCIP_Condition_Failed;
END_TRANSITION
STEP CIP4_ConditionFailed_02:
END_STEP
TRANSITION FROM CIP4_ConditionFailed_02 TO StartPump_CIP4_02
    := TRUE;
END_TRANSITION
TRANSITION FROM (Disinfct_Conc_Client_Done, Condition_CIP4_Client) TO Fill_For_MixProof_CIP4
    := bClientTypeIs_Tank AND NOT bSprinkler;
END_TRANSITION
STEP Fill_For_MixProof_CIP4:
    _aFill_For_MixProof_CIP4_entry(P1);  // entry action
    _aFill_For_MixProof_CIP4_active(N);  // step action
END_STEP
TRANSITION FROM Fill_For_MixProof_CIP4 TO Tank_MixProof_Clean_CIP4
    := bStepDone;
END_TRANSITION
STEP Tank_MixProof_Clean_CIP4:
    _aTank_MixProof_Clean_CIP4_entry(P1);  // entry action
    _aTank_MixProof_Clean_CIP4_active(N);  // step action
END_STEP
TRANSITION FROM Tank_MixProof_Clean_CIP4 TO Tank_LowLevel_CIP4_02
    := bStepDone;
END_TRANSITION
STEP Tank_LowLevel_CIP4_02:
    _aTank_LowLevel_CIP4_02_entry(P1);  // entry action
    _aTank_LowLevel_CIP4_02_active(N);  // step action
END_STEP
TRANSITION FROM Tank_LowLevel_CIP4_02 TO CIP4_Flow_Sprincler
    := bStepDone;
END_TRANSITION
STEP CIP4_Flow_Sprincler:
    _aCIP4_Flow_Sprincler_entry(P1);  // entry action
    _aCIP4_Flow_Sprincler_active(N);  // step action
END_STEP
TRANSITION FROM CIP4_Flow_Sprincler TO CIP4_Conn_Sprinkler
    := bStepDone;
END_TRANSITION
STEP CIP4_Conn_Sprinkler:
    _aCIP4_Conn_Sprinkler_entry(P1);  // entry action
    _aCIP4_Conn_Sprinkler_active(N);  // step action
END_STEP
TRANSITION FROM CIP4_Conn_Sprinkler TO StartPump_CIP4_02
    := bStepDone;
END_TRANSITION
TRANSITION FROM (Disinfct_Conc_Client_Done, Condition_CIP4_Client) TO CIP4_If_ClientIsTank
    := TRUE;
END_TRANSITION
STEP CIP4_If_ClientIsTank:
    _aCIP4_If_ClientIsTank_active(N);  // step action
END_STEP
TRANSITION FROM CIP4_If_ClientIsTank TO StopPump_CIP4_02
    := bStepDone;
END_TRANSITION
STEP StopPump_CIP4_02:  // min time T#2s
    _aStopPump_CIP4_02_entry(P1);  // entry action
END_STEP
TRANSITION FROM StopPump_CIP4_02 TO StopPump_CIP4_03
    := TRUE;
END_TRANSITION
TRANSITION FROM CIP4_If_ClientIsTank TO StopPump_CIP4_03
    := TRUE;
END_TRANSITION
STEP StopPump_CIP4_03:
    _aStopPump_CIP4_03_entry(P1);  // entry action
END_STEP
TRANSITION FROM StopPump_CIP4_03 TO Tank_LowLevel_CIP4_01
    := TRUE;
END_TRANSITION
STEP Tank_LowLevel_CIP4_01:
    _aTank_LowLevel_CIP4_01_active(N);  // step action
END_STEP
TRANSITION FROM Tank_LowLevel_CIP4_01 TO CIP4_Done
    := bStepDone;
END_TRANSITION
TRANSITION FROM Client_Check_CIP4 TO CIP4_Done
    := eReq.eClient=E_CIP_Usage.eLocal;
END_TRANSITION
STEP CIP4_Done:  // min time T#2s
    _aCIP4_Done_entry(P1);  // entry action
END_STEP
TRANSITION FROM CIP4_Done TO End_Check
    := TRUE;
END_TRANSITION
TRANSITION FROM ClientReference_IsValid TO Fill_Water_T94
    := eRun=E_CIP_Source.eT94_Water;
END_TRANSITION
// macro Water begins
STEP Fill_Water_T94:
    _aFill_Water_T94_entry(P1);  // entry action
    _aFill_Water_T94_active(N);  // step action
END_STEP
TRANSITION FROM Fill_Water_T94 TO Fill_Water_T94_Done
    := bStepDone;
END_TRANSITION
STEP Fill_Water_T94_Done:
    _aFill_Water_T94_Done_entry(P1);  // entry action
    _aFill_Water_T94_Done_active(N);  // step action
END_STEP
TRANSITION FROM Fill_Water_T94_Done TO Client_Check_CIP35
    := bStepDone;
END_TRANSITION
STEP Client_Check_CIP35:
END_STEP
TRANSITION FROM Client_Check_CIP35 TO Connect_CIP35
    := TRUE;
END_TRANSITION
STEP Connect_CIP35:
    _aConnect_CIP35_entry(P1);  // entry action
    _aConnect_CIP35_active(N);  // step action
END_STEP
TRANSITION FROM Connect_CIP35 TO StartPump_CIP35
    := bStepDone;
END_TRANSITION
STEP StartPump_CIP35:  // min time T#3s
    _aStartPump_CIP35_entry(P1);  // entry action
    _aStartPump_CIP35_active(N);  // step action
END_STEP
TRANSITION FROM StartPump_CIP35 TO CIP35_Collect
    := bStepDone;
END_TRANSITION
STEP CIP35_Collect:  // min time T#5s
    _aCIP35_Collect_entry(P1);  // entry action
    _aCIP35_Collect_active(N);  // step action
END_STEP
TRANSITION FROM CIP35_Collect TO CIP35_Drain
    := bStepDone;
END_TRANSITION
STEP CIP35_Drain:  // min time T#5s
    _aCIP35_Drain_entry(P1);  // entry action
    _aCIP35_Drain_active(N);  // step action
END_STEP
TRANSITION FROM CIP35_Drain TO Connect_CIP35_R_Water
    := bStepDone;
END_TRANSITION
STEP Connect_CIP35_R_Water:  // min time T#5s
    _aConnect_CIP35_R_Water_entry(P1);  // entry action
    _aConnect_CIP35_R_Water_active(N);  // step action
END_STEP
TRANSITION FROM Connect_CIP35_R_Water TO ReadyToCondition_Count
    := bStepDone;
END_TRANSITION
STEP ReadyToCondition_Count:
    _aReadyToCondition_Count_entry(P1);  // entry action
    _aReadyToCondition_Count_active(N);  // step action
END_STEP
TRANSITION FROM ReadyToCondition_Count TO Condition_CIP35_Client
    := TRUE;
END_TRANSITION
STEP Condition_CIP35_Client:
    _aCondition_CIP35_Client_entry(P1);  // entry action
    _aCondition_CIP35_Client_active(N);  // step action
    _aCondition_CIP35_Client_exit(P0);  // exit action
END_STEP
TRANSITION FROM Condition_CIP35_Client TO Sprinkler_Request_CIP35
    := bCIP_Condition_Done;
END_TRANSITION
STEP Sprinkler_Request_CIP35:
    _aSprinkler_Request_CIP35_active(N);  // step action
END_STEP
TRANSITION FROM Sprinkler_Request_CIP35 TO StopPump_CIP35_01
    := bStepDone;
END_TRANSITION
STEP StopPump_CIP35_01:
    _aStopPump_CIP35_01_entry(P1);  // entry action
END_STEP
TRANSITION FROM StopPump_CIP35_01 TO Tank_LowLevel_CIP35_01
    := TRUE;
END_TRANSITION
TRANSITION FROM Sprinkler_Request_CIP35 TO Tank_LowLevel_CIP35_02
    := TRUE;
END_TRANSITION
STEP Tank_LowLevel_CIP35_02:
    _aTank_LowLevel_CIP35_02_entry(P1);  // entry action
    _aTank_LowLevel_CIP35_02_active(N);  // step action
END_STEP
TRANSITION FROM Tank_LowLevel_CIP35_02 TO CIP35_Conn_Sprinkler
    := bStepDone;
END_TRANSITION
STEP CIP35_Conn_Sprinkler:
    _aCIP35_Conn_Sprinkler_entry(P1);  // entry action
    _aCIP35_Conn_Sprinkler_active(N);  // step action
END_STEP
TRANSITION FROM CIP35_Conn_Sprinkler TO ReadyToCondition_Count
    := bStepDone;
END_TRANSITION
TRANSITION FROM Condition_CIP35_Client TO StopPump_CIP35_02
    := bCIP_Condition_Failed;
END_TRANSITION
STEP StopPump_CIP35_02:
    _aStopPump_CIP35_02_entry(P1);  // entry action
END_STEP
TRANSITION FROM StopPump_CIP35_02 TO ReFill_Water_T94
    := TRUE;
END_TRANSITION
STEP ReFill_Water_T94:
    _aReFill_Water_T94_active(N);  // step action
END_STEP
TRANSITION FROM ReFill_Water_T94 TO Condition_CIP35_Client
    := bStepDone;
END_TRANSITION
STEP Tank_LowLevel_CIP35_01:
    _aTank_LowLevel_CIP35_01_active(N);  // step action
END_STEP
TRANSITION FROM Tank_LowLevel_CIP35_01 TO CIP35_Done
    := bStepDone;
END_TRANSITION
STEP CIP35_Done:  // min time T#2s
    _aCIP35_Done_entry(P1);  // entry action
END_STEP
TRANSITION FROM CIP35_Done TO End_Check
    := TRUE;
END_TRANSITION
STEP End_Check:
    _aEnd_Check_active(N);  // step action
END_STEP
TRANSITION FROM End_Check TO Disconnect_n_Drain_CIP_Client
    := bStepDone;
END_TRANSITION
TRANSITION FROM End_Check TO Get_Client
    := TRUE;
END_TRANSITION
STEP Disconnect_n_Drain_CIP_Client:
    _aDisconnect_n_Drain_CIP_Client_entry(P1);  // entry action
    _aDisconnect_n_Drain_CIP_Client_active(N);  // step action
END_STEP
TRANSITION FROM Disconnect_n_Drain_CIP_Client TO Done
    := bStepDone;
END_TRANSITION
STEP Done:  // min time T#0.1s
    _aDone_entry(P1);  // entry action
END_STEP
TRANSITION FROM Done TO Disconnect_Old_Client
    := TRUE;
END_TRANSITION
// branch label Branch28_act_Oper
// branch label Branch29_act_Oper
// branch label Branch27_act_Oper
// branch label Branch26_act_Oper
// branch label Branch0_act_Oper
// branch label Branch11_act_Oper
// branch label Branch10_act_Oper
// branch label Branch15_act_Oper
// branch label Branch14_act_Oper
// branch label Branch10_act_Oper_2
// branch label Branch23_act_Oper
// branch label Branch12_act_Oper
// branch label Branch9_act_Oper
// branch label Branch17_act_Oper
// branch label Branch18_act_Oper
// branch label Branch19_act_Oper
// branch label Branch24_act_Oper
// branch label Branch20_act_Oper
// branch label Branch8_act_Oper
// branch label Branch2_act_Oper
// branch label Branch3_act_Oper
END_ACTION

ACTION act_ReqBuffer:
rtPosMoveHMI_Up(Q=>);
IF rtPosMoveHMI_Up.Q THEN;
	m_PosMove_Up_HMI();
END_IF
rtPosMoveHMI_Down(Q=>);
IF rtPosMoveHMI_Down.Q THEN;
	m_PosMove_Down_HMI();
END_IF
rtPosDeleteHMI(Q=>);
IF rtPosDeleteHMI.Q THEN;
	m_PosDelete_HMI();
END_IF
rtPosDeleteAllHMI(Q=>);
IF rtPosDeleteAllHMI.Q THEN;
	m_PosDeleteAll_HMI();
END_IF

rtReqLocalCIP_Full_HMI(Q=>);
IF rtReqLocalCIP_Full_HMI.Q THEN;
	eReqLocal.eClient:=E_CIP_Usage.eLocal;
	eReqLocal.eType:=E_CIP_Type.Full;
	m_TakePosInCIPBuffer(stCIP_Request:=eReqLocal);
END_IF

rtReqLocalCIP_Detergent_HMI(Q=>);
IF rtReqLocalCIP_Detergent_HMI.Q THEN;
	eReqLocal.eClient:=E_CIP_Usage.eLocal;
	eReqLocal.eType:=E_CIP_Type.Detergent;
	m_TakePosInCIPBuffer(stCIP_Request:=eReqLocal);
END_IF

rtReqCleanEmpty_HMI(Q=>);
IF rtReqCleanEmpty_HMI.Q THEN;
	m_CleanEmpty_Spaces();
END_IF
END_ACTION

ACTION act_Run:
//Client error: ALARM from Siemens. Only marks the step, the reaction is in FB_CIP_Siemens
IF eReq.eClient=E_CIP_Usage.eExternal THEN;
	IF g_Anybus.fbAnybus.stIn.bAlarm AND SFCCurrentStep<>'Ready' THEN;
		m_Set_LastStepBeforeError();
		sError_Message:='Client Error';
		//mResetCycle();
	END_IF
END_IF
END_ACTION

ACTION act_SprinklerCondition:


	IF TRUE
	AND eCIP_State>=E_Element_State_Long.eCIP_1_Rinzed 
	AND eCIP_State<=E_Element_State_Long.eCIP_2_Deterged 
	THEN;
		IF NOT bSprinkler THEN // Pipe
			tConditionTime	:=st_CIP_Param.t_ConditionDetergent;
			fFlowRate		:=st_CIP_Param.r_Flow_Pipe;
		ELSE // Sprinkler
			tConditionTime	:=st_CIP_Param.t_ConditionDetergent_Sprinkler;
			fFlowRate		:=st_CIP_Param.r_Flow_Sprinkler;
		END_IF	
		//rVolume_Collect :=st_CIP_Param.r_Volume_Collect_Detergent;
		//rVolume_Drain	:=st_CIP_Param.r_Volume_Drain_Detergent;
		//rVolume_Recycle	:=st_CIP_Param.r_Volume_Recycle_Detergent;
		
	ELSIF TRUE
	AND eCIP_State>=E_Element_State_Long.eCIP_3_Deterged_Clean 
	AND eCIP_State<=E_Element_State_Long.eCIP_4_Sanitized 
	THEN;
		IF NOT bSprinkler THEN // Pipe
			tConditionTime	:=st_CIP_Param.t_ConditionDisInfection;
			fFlowRate		:=st_CIP_Param.r_Flow_Pipe;
		ELSE // Sprinkler
			tConditionTime	:=st_CIP_Param.t_ConditionDisInfection_Sprinkler;
			fFlowRate		:=st_CIP_Param.r_Flow_Sprinkler;
		END_IF	
		//rVolume_Collect :=st_CIP_Param.r_Volume_Collect_DisInfection;
		//rVolume_Drain	:=st_CIP_Param.r_Volume_Drain_DisInfection;
		//rVolume_Recycle	:=st_CIP_Param.r_Volume_Recycle_DisInfection;
	END_IF
END_ACTION

METHOD m_Set_CIP_State : BOOL
VAR_INPUT
	eState	: E_Element_State_Long;
END_VAR
//CIP stages only move forward (eNotClean restarts)
IF (eState>eCIP_State
OR eState=E_Element_State_Long.eNotClean)
AND eState<=E_Element_State_Long.eProduction
THEN;
	eCIP_State:=eState;
	m_Set_CIP_State:=TRUE;
END_IF
END_METHOD

METHOD m_DashState_NotAvailable : BOOL
VAR_INPUT
	stage: E_CIP_DashStage_List;
END_VAR
//Client and sprinkler stages do not exist in the local CIP
CASE stage OF
	E_CIP_DashStage_List.e01_CIP1_Client_Drain_Product_Rest_Pipe,
	E_CIP_DashStage_List.e02_CIP1_Client_Drain_Product_Rest_Sprinkler,
	E_CIP_DashStage_List.e05_CIP2_Client_Detergent_Fill,
	E_CIP_DashStage_List.e06_CIP2_Client_Detergent_Condition_Pipe,
	E_CIP_DashStage_List.e07_CIP2_Client_Detergent_Condition_Sprinkler,
	E_CIP_DashStage_List.e11_CIP3_Detergent_Clean_Sprinkler,
	E_CIP_DashStage_List.e14_CIP4_Client_DisInfection_Fill,
	E_CIP_DashStage_List.e15_CIP4_Client_DisInfection_Condition_Pipe,
	E_CIP_DashStage_List.e16_CIP4_Client_DisInfection_Condition_Sprinkler,
	E_CIP_DashStage_List.e20_CIP5_DisInfection_Clean_Sprinkler:;
		m_DashState_NotAvailable:=TRUE;
ELSE;
		m_DashState_NotAvailable:=FALSE;
END_CASE
END_METHOD

METHOD m_Check_ProductionTank_Low_Level : BOOL
VAR_INPUT
END_VAR
//The client level is on the plant side: Tank waits for CLIENT EMPTY, as senLL before, Pipe passes
tonTankLowLevel.IN:=g_Anybus.fbAnybus.stIn.bClientEmpty;
tonTankLowLevel(PT:=T#2S);
IF bClientTypeIs_Tank
AND tonTankLowLevel.Q
THEN;
	m_Check_ProductionTank_Low_Level:=TRUE;
ELSIF NOT bClientTypeIs_Tank
THEN;
	m_Check_ProductionTank_Low_Level:=TRUE;
ELSE;
	m_Check_ProductionTank_Low_Level:=FALSE;
END_IF
END_METHOD

METHOD m_CleanEmpty_Spaces : BOOL
VAR_INPUT
END_VAR

VAR
	i: INT;
	j: INT;
	stCIP_Request_Empty: ST_CIP_Request;
END_VAR
FOR i:=0 TO 9 DO
	IF i<>0 OR NOT bRun THEN;
		IF arCIP_RequestBufer[i].eClient=E_CIP_Usage.eNotInUse THEN;
			FOR j:=i+1 TO 9 DO
				IF arCIP_RequestBufer[j].eClient<>E_CIP_Usage.eNotInUse THEN;
					arCIP_RequestBufer[i]:=arCIP_RequestBufer[j];
					arCIP_RequestBufer[j]:=stCIP_Request_Empty;
					EXIT;
				END_IF
			END_FOR
		END_IF		
	END_IF
END_FOR
END_METHOD

METHOD m_ClientTank_IsEmpty : BOOL
VAR_INPUT
END_VAR
IF __ISVALIDREF(ref_lvlTank_Client) 
AND bClientTypeIs_Tank
THEN;
	m_ClientTank_IsEmpty:=ref_lvlTank_Client.e_state=E_Tank_Level.eEmpty;
ELSE;
	m_ClientTank_IsEmpty:=TRUE;
END_IF
END_METHOD

METHOD m_ClientTank_Level_IsHigher_Then : BOOL
VAR_INPUT
	min_Level: REAL:=150.0;
END_VAR
IF __ISVALIDREF(ref_lvlTank_Client) 
AND bClientTypeIs_Tank
THEN;
	m_ClientTank_Level_IsHigher_Then:=ref_lvlTank_Client.rTankLevel>=min_Level;
ELSE;
	m_ClientTank_Level_IsHigher_Then:=FALSE;
END_IF
END_METHOD

METHOD m_DashState_activate : BOOL
VAR_INPUT
	stage		: E_CIP_DashStage_List;
END_VAR
	IF arCIP_DashStage_list[stage] = E_CIP_DashStage.eCIPStage_ToBeDone THEN;
		arCIP_DashStage_list[stage]:=E_CIP_DashStage.eCIPStage_Active;
		eCIP_DashStage_actual:=stage;
		sCIP_DashStage_actual:=TO_STRING(eCIP_DashStage_actual);	
		RETURN;
	END_IF

(*
FOR stage:=m_DashState_from() TO m_DashState_to() DO
	IF arCIP_DashStage_list[stage] = E_CIP_DashStage.eCIPStage_ToBeDone THEN;
		arCIP_DashStage_list[stage]:=E_CIP_DashStage.eCIPStage_Active;
		eCIP_DashStage_actual:=stage;
		sCIP_DashStage_actual:=TO_STRING(eCIP_DashStage_actual);	
		RETURN;
	END_IF
END_FOR
*)
END_METHOD

METHOD m_DashState_done : BOOL
VAR_INPUT
	stage	: E_CIP_DashStage_List;
END_VAR
IF arCIP_DashStage_list[stage] = E_CIP_DashStage.eCIPStage_Active THEN;
	arCIP_DashStage_list[stage]:=E_CIP_DashStage.eCIPStage_Done;
	RETURN;
END_IF

(*
FOR stage:=m_DashState_from() TO m_DashState_to() DO
	IF arCIP_DashStage_list[stage] = E_CIP_DashStage.eCIPStage_Active THEN;
		arCIP_DashStage_list[stage]:=E_CIP_DashStage.eCIPStage_Done;
		RETURN;
	END_IF
END_FOR
*)
END_METHOD

METHOD m_DashState_from : E_CIP_DashStage_List
VAR
	eActCIP_State	: E_Element_State_Long;
END_VAR
eActCIP_State:=eCIP_State;

CASE eActCIP_State OF
	E_Element_State_Long.eNotClean:;
		m_DashState_from:=E_CIP_DashStage_List.e01_CIP1_Client_Drain_Product_Rest_Pipe;	
		
	E_Element_State_Long.eCIP_1_Rinzed:;
		m_DashState_from:=E_CIP_DashStage_List.e03_CIP2_Local_Detergent_Fill;	
	
	E_Element_State_Long.eCIP_2_Deterged:;
		m_DashState_from:=E_CIP_DashStage_List.e08_CIP3_Detergent_Collect;	
	
	E_Element_State_Long.eCIP_3_Deterged_Clean:;
		m_DashState_from:=E_CIP_DashStage_List.e12_CIP4_Local_DisInfection_Fill;	
	
	E_Element_State_Long.eCIP_4_Sanitized:;
		m_DashState_from:=E_CIP_DashStage_List.e17_CIP5_DisInfection_Collect;	
	
ELSE;
	//???
		m_DashState_from:=E_CIP_DashStage_List.eLast;
END_CASE
END_METHOD

METHOD m_DashState_Get_ToBeDone_List : BOOL
VAR
	//eActCIP_State	: E_Element_State_Long;
	//eCIP_req		: ST_CIP_Request;	
	stage			: E_CIP_DashStage_List;
END_VAR
//eCIP_req:=eReq;

//init
FOR stage:=E_CIP_DashStage_List.e00_NotSelected TO E_CIP_DashStage_List.eLast DO
	arCIP_DashStage_list[stage]:=E_CIP_DashStage.eCIPStage_NotAvalable;
END_FOR

//Start done condition stages
FOR stage:=E_CIP_DashStage_List.e00_NotSelected TO m_DashState_from()-1 DO
	IF m_DashState_Sprinkler(stage:=stage) THEN;
		IF bClientTypeIs_Tank THEN;
			arCIP_DashStage_list[stage]:=E_CIP_DashStage.eCIPStage_Done;
		ELSE;
			arCIP_DashStage_list[stage]:=E_CIP_DashStage.eCIPStage_NotAvalable;
		END_IF
	ELSE;
		arCIP_DashStage_list[stage]:=E_CIP_DashStage.eCIPStage_Done;
	END_IF
END_FOR

// Request conditions
FOR stage:=m_DashState_from() TO m_DashState_to() DO
	IF m_DashState_Sprinkler(stage:=stage) THEN;
		IF bClientTypeIs_Tank THEN;
			arCIP_DashStage_list[stage]:=E_CIP_DashStage.eCIPStage_ToBeDone;
		ELSE;
			arCIP_DashStage_list[stage]:=E_CIP_DashStage.eCIPStage_NotAvalable;
		END_IF
	ELSE;
		arCIP_DashStage_list[stage]:=E_CIP_DashStage.eCIPStage_ToBeDone;
	END_IF
END_FOR

//Do not requested 
FOR stage:=m_DashState_to()+1 TO E_CIP_DashStage_List.eLast DO
	IF m_DashState_Sprinkler(stage:=stage) THEN;
		IF bClientTypeIs_Tank THEN;
			arCIP_DashStage_list[stage]:=E_CIP_DashStage.eCIPStage_NotInUse;
		ELSE;
			arCIP_DashStage_list[stage]:=E_CIP_DashStage.eCIPStage_NotAvalable;
		END_IF
	ELSE;
		arCIP_DashStage_list[stage]:=E_CIP_DashStage.eCIPStage_NotInUse;
	END_IF
END_FOR
END_METHOD

METHOD m_DashState_Sprinkler : BOOL
VAR_INPUT
	stage: E_CIP_DashStage_List;
END_VAR
CASE stage OF 
	E_CIP_DashStage_List.e02_CIP1_Client_Drain_Product_Rest_Sprinkler,
	E_CIP_DashStage_List.e07_CIP2_Client_Detergent_Condition_Sprinkler,
	E_CIP_DashStage_List.e11_CIP3_Detergent_Clean_Sprinkler,
	E_CIP_DashStage_List.e16_CIP4_Client_DisInfection_Condition_Sprinkler,
	E_CIP_DashStage_List.e20_CIP5_DisInfection_Clean_Sprinkler:;
		m_DashState_Sprinkler:=TRUE;
ELSE;
		m_DashState_Sprinkler:=FALSE;
END_CASE
END_METHOD

METHOD m_DashState_to : E_CIP_DashStage_List
VAR
	eCIP_req		: ST_CIP_Request;
END_VAR
eCIP_req:=eReq;

CASE eCIP_req.eType OF
	E_CIP_Type.R_Water:;
		m_DashState_to:=E_CIP_DashStage_List.e02_CIP1_Client_Drain_Product_Rest_Sprinkler;
		
	E_CIP_Type.Detergent:;
		m_DashState_to:=E_CIP_DashStage_List.e11_CIP3_Detergent_Clean_Sprinkler;
	
	E_CIP_Type.Full:;
		m_DashState_to:=E_CIP_DashStage_List.e20_CIP5_DisInfection_Clean_Sprinkler;

ELSE;
	//???
		m_DashState_to:=E_CIP_DashStage_List.eLast;	
END_CASE
END_METHOD

METHOD m_DashState_ToString_convertion : BOOL
VAR_INPUT
END_VAR

VAR
	eDashboard_CIP_State: E_CIP_DashStage_List:=E_CIP_DashStage_List.eLast;
END_VAR
FOR eDashboard_CIP_State:=0 TO E_CIP_DashStage_List.eLast DO
	//g_HMI.arCIP_DashStage_list[eDashboard_CIP_State]:=E_CIP_DashStage.eCIPStage_NotInUse;
	g_HMI.arCIP_DashStage_string[eDashboard_CIP_State]:=TO_STRING(eDashboard_CIP_State);
END_FOR
END_METHOD

METHOD m_MeasureTimeToHMI : TIME
VAR_INPUT
END_VAR
IF SFCCurrentStep='measureDelay_CIP2_1' THEN;
	m_MeasureTimeToHMI:=measureDelay_CIP2_1.t;
	
ELSIF SFCCurrentStep='measureDelay_CIP2_2' THEN;
	m_MeasureTimeToHMI:=measureDelay_CIP2_2.t;
	
ELSIF SFCCurrentStep='measureDelay_CIP4_1' THEN;
	m_MeasureTimeToHMI:=measureDelay_CIP4_1.t;
	
ELSIF SFCCurrentStep='measureDelay_CIP4_2' THEN;
	m_MeasureTimeToHMI:=measureDelay_CIP4_2.t;

ELSE;
	m_MeasureTimeToHMI:=T#0S;
END_IF
END_METHOD

METHOD m_OverFlowCorrect : REAL
VAR_INPUT
	rTc		:	REAL	;//Target concentration
	rAv		:	REAL	;//Actual volume
	rAc		:	REAL	;//Actual concentration
END_VAR
//Calculating the additional valume of fresh water to dalute the concentration
IF rTc=0 THEN;
	m_OverFlowCorrect:=0;
ELSE;
	m_OverFlowCorrect:=((rAv*rAc/100)/(rTc/100))-(rAv*rAc/100)-rAv+(rAv*rAc/100);
END_IF
END_METHOD

METHOD m_PosDelete_HMI : BOOL
VAR_INPUT
END_VAR
VAR
	stCIP_Request_Empty: ST_CIP_Request;
END_VAR
IF iPosSelect_HMI>=0 AND iPosSelect_HMI<9 THEN;
	IF iPosSelect_HMI<>0 OR NOT bRun THEN;
		arCIP_RequestBufer[iPosSelect_HMI]:=stCIP_Request_Empty;
	END_IF		
END_IF
END_METHOD

METHOD m_PosDeleteAll_HMI : BOOL
VAR_INPUT
END_VAR
VAR
	stCIP_Request_Empty: ST_CIP_Request;
	i: INT;
END_VAR

FOR i:=0 TO 9 DO
	IF i<>0 OR NOT bRun THEN;
		arCIP_RequestBufer[i]:=stCIP_Request_Empty;
	END_IF	
END_FOR
END_METHOD

METHOD m_PosMove_Down_HMI : BOOL
VAR_INPUT
END_VAR
VAR
	stCIP_Request_Temp: ST_CIP_Request;
	i: INT;
END_VAR
IF iPosSelect_HMI>=0 AND iPosSelect_HMI<9 THEN;
	IF iPosSelect_HMI<>0 OR NOT bRun THEN;		
			IF ((arCIP_RequestBufer[iPosSelect_HMI].eType=E_CIP_Type.R_Water 
				AND (arCIP_RequestBufer[iPosSelect_HMI+1].eType=E_CIP_Type.Detergent 
				OR arCIP_RequestBufer[iPosSelect_HMI+1].eType=E_CIP_Type.Full)) 
			OR (arCIP_RequestBufer[iPosSelect_HMI].eType=E_CIP_Type.Detergent 				
				AND arCIP_RequestBufer[iPosSelect_HMI+1].eType=E_CIP_Type.Full))
			AND (arCIP_RequestBufer[iPosSelect_HMI+1].eClient=arCIP_RequestBufer[iPosSelect_HMI].eClient) 
			THEN
				;
			ELSE
				stCIP_Request_Temp:=arCIP_RequestBufer[iPosSelect_HMI+1];
				arCIP_RequestBufer[iPosSelect_HMI+1]:=arCIP_RequestBufer[iPosSelect_HMI];
				arCIP_RequestBufer[iPosSelect_HMI]:=stCIP_Request_Temp;
				iPosSelect_HMI:=iPosSelect_HMI+1;	
			END_IF	
	END_IF
END_IF
END_METHOD

METHOD m_PosMove_Up_HMI : BOOL
VAR_INPUT
END_VAR
VAR
	stCIP_Request_Temp: ST_CIP_Request;
	i: INT;
	m: bool;
END_VAR
IF iPosSelect_HMI>0 AND iPosSelect_HMI<=9 THEN;
	IF iPosSelect_HMI<>1 OR NOT bRun THEN;			
			IF ((arCIP_RequestBufer[iPosSelect_HMI].eType=e_cip_type.Full 
				AND (arCIP_RequestBufer[iPosSelect_HMI-1].eType=E_CIP_Type.Detergent 
				OR arCIP_RequestBufer[iPosSelect_HMI-1].eType=E_CIP_Type.R_Water)) 
			OR (arCIP_RequestBufer[iPosSelect_HMI].eType=E_CIP_Type.Detergent 
				AND arCIP_RequestBufer[iPosSelect_HMI-1].eType=E_CIP_Type.R_Water))
			AND (arCIP_RequestBufer[iPosSelect_HMI-1].eClient=arCIP_RequestBufer[iPosSelect_HMI].eClient) 
			THEN
				;
			ELSE
				stCIP_Request_Temp:=arCIP_RequestBufer[iPosSelect_HMI-1];
				arCIP_RequestBufer[iPosSelect_HMI-1]:=arCIP_RequestBufer[iPosSelect_HMI];
				arCIP_RequestBufer[iPosSelect_HMI]:=stCIP_Request_Temp;
				iPosSelect_HMI:=iPosSelect_HMI-1;
			END_IF	
	END_IF
END_IF
END_METHOD

METHOD m_Set_SFCFlags_Reference : BOOL
//Set reference to SFC flags

refSFC.SFCInit REF= SFCInit;
refSFC.SFCReset REF= SFCReset;
refSFC.SFCError REF= SFCError;
refSFC.SFCEnableLimit REF= SFCEnableLimit;
refSFC.SFCErrorStep REF= SFCErrorStep;
refSFC.SFCErrorPOU REF= SFCErrorPOU;
refSFC.SFCQuitError REF= SFCQuitError;
refSFC.SFCPause REF= SFCPause;
refSFC.SFCTrans REF= SFCTrans;
refSFC.SFCCurrentStep REF= SFCCurrentStep;
refSFC.SFCTip REF= SFCTip;
refSFC.SFCTipMode REF= SFCTipMode;

// Cycle handle for SFC
m_SFC_Handle();

m_Set_Mode_Reference(inMoedeZone:=E_ModeZone.eCIP);
END_METHOD

METHOD m_TakePosInCIPBuffer : BOOL
VAR_INPUT
	stCIP_Request: ST_CIP_Request;
END_VAR

VAR
	i: INT;
	m: bool;	
END_VAR
//Old client checks (production, state, duplicate), not used for eExternal, fbElement is removed
(*
IF stCIP_Request.eClient<>E_CIP_Usage.eNotInUse
AND stCIP_Request.eType<>E_CIP_Type.NotSelected
AND g_data.fbElement[stCIP_Request.eClient].ProdStatus<>E_Prod_Status.Active
AND g_data.fbElement[stCIP_Request.eClient].eState_Long>E_Element_State_Long.eStandby 
AND ((stCIP_Request.eType=E_CIP_Type.R_Water AND g_data.fbElement[stCIP_Request.eClient].eState_Long<E_Element_State_Long.eCIP_1_Rinzed)
	OR (stCIP_Request.eType=E_CIP_Type.Detergent AND g_data.fbElement[stCIP_Request.eClient].eState_Long<E_Element_State_Long.eCIP_3_Deterged_Clean)
	OR (stCIP_Request.eType=E_CIP_Type.Full AND g_data.fbElement[stCIP_Request.eClient].eState_Long<E_Element_State_Long.eCIP_5_Done))

THEN
	FOR i:=0 TO 9 DO
		IF arCIP_RequestBufer[i].eClient=stCIP_Request.eClient 
			AND arCIP_RequestBufer[i].eType>=stCIP_Request.eType 
		THEN 	
				m:=FALSE;
				EXIT;
			ELSE
				m:=TRUE;
		END_IF
	END_FOR	
	IF m=TRUE THEN
		FOR i:=0 TO 9 DO
			IF arCIP_RequestBufer[i].eClient=E_CIP_Usage.eNotInUse 
			THEN;
				arCIP_RequestBufer[i]:=stCIP_Request;
				m:=FALSE;
				EXIT;
			END_IF
		END_FOR	
	END_IF
ELSIF stCIP_Request.eClient=E_CIP_Usage.eLocal
AND stCIP_Request.eType<>E_CIP_Type.NotSelected
THEN;
		FOR i:=0 TO 9 DO
			IF arCIP_RequestBufer[i].eClient=E_CIP_Usage.eNotInUse 
			THEN;
				arCIP_RequestBufer[i]:=stCIP_Request;
				m:=FALSE;
				EXIT;
			END_IF
		END_FOR		
END_IF
*)
//R_Water is not a valid local request
IF (stCIP_Request.eClient=E_CIP_Usage.eLocal
	AND (stCIP_Request.eType=E_CIP_Type.Detergent OR stCIP_Request.eType=E_CIP_Type.Full))
OR (stCIP_Request.eClient=E_CIP_Usage.eExternal
	AND stCIP_Request.eType<>E_CIP_Type.NotSelected)
THEN;
		FOR i:=0 TO 9 DO
			IF arCIP_RequestBufer[i].eClient=E_CIP_Usage.eNotInUse
			THEN;
				arCIP_RequestBufer[i]:=stCIP_Request;
				m:=FALSE;
				EXIT;
			END_IF
		END_FOR
END_IF
END_METHOD

METHOD mFillWater : BOOL
VAR_INPUT
END_VAR

VAR
	reqVolume: REAL;	
	valve : E_Pis_Name;;
	actLevel: REAL;
	fillCondition: BOOL;	
	
END_VAR
IF TRUE 
AND fbPis.m_CheckByRecipe(stPis:=stPis_FillWater_T91, req:=E_Piston_Recipe_State.Release)
AND fbPis.m_CheckByRecipe(stPis:=stPis_FillWater_T92, req:=E_Piston_Recipe_State.Release)
AND fbPis.m_CheckByRecipe(stPis:=stPis_FillWater_T93, req:=E_Piston_Recipe_State.Release)
AND bStateSafe
AND MAIN.bTemp_Water_Overweight_check
THEN;
	fillCondition:=TRUE;
ELSE;
	fillCondition:=FALSE;
END_IF

reqVolume:=st_CIP_Param.r_Tank94_Volume;
IF g_Data.arr_CIP_Recipe[nLocalRecipe].r_Tank94_Volume>reqVolume THEN;
	reqVolume:=g_Data.arr_CIP_Recipe[nLocalRecipe].r_Tank94_Volume;
END_IF

fbHysteresisFillT94(
	fIn:= lvlTank_T94.rTankLevel, 
	fHigh:= reqVolume, 
	fLow:= reqVolume-50.0, 
	iDigitsAfterDot:= 1, 
	bOut=> );

IF eMode<>E_CIP_Mode.eOff THEN;
	IF fbPis.m_CheckByRecipe(stPis:=stPis_FillWater_T94, req:=E_Piston_Recipe_State.Act) 
	AND (NOT fbHysteresisFillT94.bOut
	OR NOT fillCondition)
	THEN;
		//stPis_FillWater_T94.req_Close:=TRUE;
		fbPis.m_SetByRecipe(stPis:=stPis_FillWater_T94, req:=E_Piston_Recipe_State.Release);
		
	ELSIF fbPis.m_CheckByRecipe(stPis:=stPis_FillWater_T94, req:=E_Piston_Recipe_State.Release) 
	AND fbHysteresisFillT94.bOut
	AND fillCondition
	THEN;
		IF NOT arrTanksSens[E_Tank_Name.T94].get_stTankLevel_OverFlow() THEN;
			fbPis.m_SetByRecipe(stPis:=stPis_FillWater_T94, req:=E_Piston_Recipe_State.Act);			
		END_IF	
	END_IF	
END_IF
	
	
(*
fbFillT94(	
		valve:= valFillWater_T94, 
		reqLevel:= reqVolume, 
		actLevel:= lvlTank_T94.rTankLevel, 
		fillCondition:= );
*)
END_METHOD

METHOD mLoadDefProcessSetPoints : BOOL
VAR_INPUT
END_VAR

	stDetergent.ToleranceHigh:=0.05;
	stDetergent.ToleravceLow:=0.05;
	stTemperature_Deterg.ToleranceHigh:=1;
	stTemperature_Deterg.ToleravceLow:=1;
	stDisInfectant.ToleranceHigh:=0.05;
	stDisInfectant.ToleravceLow:=0.05;
	stTemperature_Dis.ToleranceHigh:=1;//0.5
	stTemperature_Dis.ToleravceLow:=1;//0.5
	stFlow1_Rate.ToleranceHigh:=10;
	stFlow1_Rate.ToleravceLow:=10;
	stFlow2_Rate.ToleranceHigh:=10;
	stFlow2_Rate.ToleravceLow:=10;
	stP1001_Pressure.ToleranceHigh:=1;
	stP1001_Pressure.ToleravceLow:=1;
END_METHOD

METHOD mProcessDeviation : REAL
VAR_INPUT
	reqValue: REAL;
	processValue: REAL;
END_VAR
mProcessDeviation:=reqValue-processValue;
END_METHOD

METHOD mVolumeMeter : BOOL
VAR_INPUT
END_VAR
delta_T91_Volume:=lvlTank_T91.rTankLevel-memo_T91_Level_start;//de
delta_T92_Volume:=lvlTank_T92.rTankLevel-memo_T92_Level_start;
delta_T93_Volume:=lvlTank_T93.rTankLevel-memo_T93_Level_start;
delta_T94_Volume:=lvlTank_T94.rTankLevel-memo_T94_Level_start;
END_METHOD

METHOD mVolumeReset_All : BOOL
VAR_INPUT
END_VAR
memo_T91_Level_start:=lvlTank_T91.rTankLevel;
memo_T92_Level_start:=lvlTank_T92.rTankLevel;
memo_T93_Level_start:=lvlTank_T93.rTankLevel;
memo_T94_Level_start:=lvlTank_T94.rTankLevel;
END_METHOD

END_FUNCTION_BLOCK

(* stored: Version 1.1.0.1, ProductVersion 3.1.4026.20
   POU FB_CIP: Id {14cc32b0-9432-4cf7-99d2-9b696d5c02b0}, SpecialFunc None
   Folder Manage: Id {8cb05385-d8fc-420c-9505-d8b2a8121243}
   Folder Meth: Id {3ff852d5-11b9-4725-a976-204de9549283}
   Folder Dashboard: Id {9e04f67f-2723-4849-a13e-a86c894f0a2f}
   Folder HMI_queue_pos: Id {5c4eceae-9a17-444f-b26e-881c006e97cc}
   Action _aCIP1_Conn_Sprinkler_active: Id {4c796a07-4449-4c49-bcc2-457b99419775}
   Action _aCIP1_Conn_Sprinkler_entry: Id {5b8727b3-8cd5-4a98-a184-e51877734957}
   Action _aCIP1_Done_entry: Id {5876c70f-a066-4ad6-a135-a5384197da92}
   Action _aCIP2_Conn_Sprinkler_active: Id {fa73b005-a258-42c6-9c70-008e2384c458}
   Action _aCIP2_Conn_Sprinkler_entry: Id {6c3ad8e1-0a21-4e23-9194-b2e6b28ff999}
   Action _aCIP2_Done_entry: Id {9a18f41c-f03b-4bca-ad35-6eeccc6aba8e}
   Action _aCIP2_Flow_Sprincler_active: Id {2abfbe97-fb20-494a-be0b-de7a5d389ef0}
   Action _aCIP2_Flow_Sprincler_entry: Id {4454f205-0cdf-4ef6-883c-72552e22abc1}
   Action _aCIP2_If_ClientIsTank_active: Id {4a9144df-9ae3-4d28-9b85-5b9ce93c547e}
   Action _aCIP4_Conn_Sprinkler_active: Id {74ae984f-0ae0-4e0b-96ce-fe160b8e69b3}
   Action _aCIP4_Conn_Sprinkler_entry: Id {2d20e61c-61b4-4d4d-a421-445dee37edfa}
   Action _aCIP4_Done_entry: Id {ea9db615-0bf9-482c-b261-eaf0de2b9036}
   Action _aCIP4_Flow_Sprincler_active: Id {852cab69-83b0-43ef-990f-f698125ebc48}
   Action _aCIP4_Flow_Sprincler_entry: Id {507a1c3c-2446-4445-99e2-6371dfdeab5d}
   Action _aCIP4_If_ClientIsTank_active: Id {e5c94bea-403b-4ee1-a03c-d5388d877ad2}
   Action _aCIP35_Collect_active: Id {245a31fa-2345-490d-951c-e73052de6876}
   Action _aCIP35_Collect_entry: Id {6daf871f-9050-473d-9190-81d975256abb}
   Action _aCIP35_Conn_Sprinkler_active: Id {e4186464-92a5-4be4-b6cb-cca91a77c405}
   Action _aCIP35_Conn_Sprinkler_entry: Id {b8e2edd9-6091-4c93-a395-b9fac0caddc7}
   Action _aCIP35_Done_entry: Id {2c90a1c0-9583-407e-b51f-9727c492c562}
   Action _aCIP35_Drain_active: Id {d7aa4e20-df54-48dd-9a3c-3664a01991e5}
   Action _aCIP35_Drain_entry: Id {048a2c59-3991-477e-82b6-2061ef66a49f}
   Action _aClient_tank_IsEmpty_active: Id {becf051e-545c-47b6-9688-7e31c59b9a42}
   Action _aClient_Validation_check_active: Id {944b4ef3-9c09-45a7-92e7-559823a6a540}
   Action _aClientReference_IsValid_entry: Id {a12df6dc-c969-4946-9c7b-d8b72cd2928a}
   Action _aCondition_CIP1_Client_active: Id {9c9aa498-c10a-4f64-a491-9b8cc01cad7d}
   Action _aCondition_CIP1_Client_entry: Id {649219db-8d44-4e51-8e61-14138dc431b7}
   Action _aCondition_CIP1_Client_exit: Id {0b2f759b-35ea-4c43-9c5b-8016affab793}
   Action _aCondition_CIP2_Client_active: Id {4c374eda-5cab-4d42-be48-b4cc4764cc7c}
   Action _aCondition_CIP2_Client_exit: Id {757d5740-8244-401c-a747-366cb0fbe409}
   Action _aCondition_CIP2_Local_active: Id {e5e07d09-44e8-4297-94d3-a998af75e5e0}
   Action _aCondition_CIP2_Local_exit: Id {3abd6e3a-fa29-4e39-83b3-0f68581fb9ea}
   Action _aCondition_CIP4_Client_active: Id {c8b10d3e-d2df-4479-877a-926158cbaf79}
   Action _aCondition_CIP4_Client_exit: Id {28991b97-1b79-4eab-99eb-3915fef0281d}
   Action _aCondition_CIP4_Local_active: Id {df016d92-2d66-4702-a496-5eb5a36fcd94}
   Action _aCondition_CIP4_Local_exit: Id {c5ddd08b-9232-4cf0-8f74-a26e6c7d4c1f}
   Action _aCondition_CIP35_Client_active: Id {bfe6d02a-b7ef-406a-9930-97a8c275e005}
   Action _aCondition_CIP35_Client_entry: Id {d3c6cb88-c31f-437c-b71e-7c943a37e052}
   Action _aCondition_CIP35_Client_exit: Id {b13fef85-6437-4f3c-bbb4-774296215049}
   Action _aConnect_CIP1_Drain_active: Id {027bf863-1ae4-4bdd-8945-394ab7bb998b}
   Action _aConnect_CIP1_Drain_entry: Id {f8896680-aaad-4c37-8e47-205e55062b9d}
   Action _aConnect_CIP2_01_active: Id {44126bcf-d2e3-4d19-8c41-62bc81f03fcf}
   Action _aConnect_CIP2_01_entry: Id {706022d5-0f64-404a-afba-3efb082d83da}
   Action _aConnect_CIP2_02_active: Id {4bc23466-f84b-4f74-9fd7-7d261847025c}
   Action _aConnect_CIP2_02_entry: Id {26108fe3-9f83-4c60-a43f-30cdb9c5ae88}
   Action _aConnect_CIP2_Drain_active: Id {cc8a26b6-3142-4ea7-a379-53edb9e4d6fd}
   Action _aConnect_CIP2_Drain_entry: Id {f852288b-60ab-4030-a5d9-399179d0fac3}
   Action _aConnect_CIP4_01_active: Id {6ad9d3b4-017f-4b24-b262-50ad8667ca02}
   Action _aConnect_CIP4_01_entry: Id {18fdbb91-79bd-4d84-b4f8-b9f91bf5c71e}
   Action _aConnect_CIP4_02_active: Id {792efcc2-564d-489b-9d68-8f14ba3ef505}
   Action _aConnect_CIP4_02_entry: Id {3d7e9a21-8eb7-46bc-aab2-fb63e0bca5ca}
   Action _aConnect_CIP4_Drain_active: Id {0d17ae16-8ab4-4fa4-adea-80b5db954086}
   Action _aConnect_CIP4_Drain_entry: Id {0ac31c05-8c73-425f-955c-b721846a3dd9}
   Action _aConnect_CIP35_active: Id {588b6467-3c69-4e91-bbae-17dceb39c081}
   Action _aConnect_CIP35_entry: Id {e2d0dcfe-cb47-41eb-a6a5-6136c5fde635}
   Action _aConnect_CIP35_R_Water_active: Id {807c7e93-dfb5-427d-b401-c9085b8404a0}
   Action _aConnect_CIP35_R_Water_entry: Id {14a8e164-fee8-4fa5-b39e-b5e01295e23f}
   Action _aDeterg_Dose_1_active: Id {adf67c15-5e80-4d92-80d5-80ed13167f81}
   Action _aDeterg_Dose_2_active: Id {409e36b4-ce3e-45aa-93de-65e556464419}
   Action _aDeterg_Overflow_1_active: Id {cd08c8a2-15e0-4912-b571-0d97b1994428}
   Action _aDeterg_Overflow_1_entry: Id {f52b8f3a-d9dc-44f3-86b4-8408e5527d40}
   Action _aDeterg_Overflow_2_active: Id {885afaf6-dc59-4f6b-8c27-9f845d09afe7}
   Action _aDeterg_Overflow_2_entry: Id {aed20db8-6bd2-40ba-bd59-a785dcee6c2b}
   Action _aDisconnect_n_Drain_CIP_Client_active: Id {0908cf68-67b7-4a91-b7fc-e2282fd9e163}
   Action _aDisconnect_n_Drain_CIP_Client_entry: Id {389c4393-cc6f-44b7-aa76-d6cd696fd6a2}
   Action _aDisconnect_Old_Client_entry: Id {0737bcf1-8ed2-4576-9f1e-32273d33eec5}
   Action _aDisinfct_Dose_1_active: Id {13f0b073-1394-4ea7-a7b7-4f151e56d9d5}
   Action _aDisinfct_Dose_2_active: Id {70662d8d-9a1e-471d-ac18-b200f397466b}
   Action _aDisinfct_Overflow_1_active: Id {4596c1cb-87de-42cb-9a79-bdfa938453a5}
   Action _aDisinfct_Overflow_1_entry: Id {2b4f5e27-bf29-490e-8560-26cd3cd60949}
   Action _aDisinfct_Overflow_2_active: Id {27431b62-dbc9-4a59-858c-5c0e54196656}
   Action _aDisinfct_Overflow_2_entry: Id {0fc6b6de-3854-4bc2-ab3c-0f51b6b56683}
   Action _aDone_entry: Id {65c51eeb-ff71-4a7b-932e-5755a43e7ba7}
   Action _aEnd_Check_active: Id {98177335-fdd1-4c16-8092-a4d30c9fc2e4}
   Action _aFill_For_MixProof_CIP2_active: Id {e817e6b9-943e-4538-ae34-690c92c75322}
   Action _aFill_For_MixProof_CIP2_entry: Id {f06ef343-5e0d-40f5-a01b-5b215dc5ed5e}
   Action _aFill_For_MixProof_CIP4_active: Id {0b721ed8-2911-4d99-9faa-f99991d07393}
   Action _aFill_For_MixProof_CIP4_entry: Id {bc672a0a-e606-4356-a465-98f1944e9811}
   Action _aFill_Solution_CIP2_active: Id {9d6ff8fa-91bd-4c22-8820-620f672402fa}
   Action _aFill_Solution_CIP4_active: Id {74e111a2-69e4-43d1-a5ee-7e24dfbfb5e1}
   Action _aFill_Solution_CIP4_entry: Id {0bc51ded-0fb2-48b2-a7f6-a093346aa47f}
   Action _aFill_Water_T91_active: Id {5095c3b6-e26a-419b-998b-d45425bd5a3c}
   Action _aFill_Water_T91_entry: Id {9e52c220-fb12-4b0d-9ba6-fd0ad192da08}
   Action _aFill_Water_T92_active: Id {24710a65-e152-4b5e-946e-ece3bbec20c5}
   Action _aFill_Water_T92_entry: Id {8d73f55e-b96a-48ae-b162-9be1fecb7a86}
   Action _aFill_Water_T93_active: Id {b2a4014f-5739-46d3-b6aa-1609eef63419}
   Action _aFill_Water_T93_Done_active: Id {b1e57830-4ca3-48e1-ba83-90b3963236c8}
   Action _aFill_Water_T93_Done_entry: Id {6d4baf80-ad8d-4a30-bf72-135be7a85309}
   Action _aFill_Water_T93_entry: Id {b00c63f0-fee4-40ed-826a-0670a2235d2b}
   Action _aFill_Water_T94_active: Id {69b06cae-7ea8-4e4a-93f0-c2b1370a9df2}
   Action _aFill_Water_T94_Done_active: Id {972d8a9c-6f90-434c-9eee-b7777733be46}
   Action _aFill_Water_T94_Done_entry: Id {287195c7-6b19-4c7c-93db-2e108a95040c}
   Action _aFill_Water_T94_entry: Id {cab8dd8a-41d7-4bc6-8864-94606c706eb3}
   Action _aFlow_Volume_Meter_active: Id {4cd929bd-0e77-4721-bfed-4c0b7b4378fd}
   Action _aGet_Client_active: Id {18e627b5-82b2-485b-93fe-c20af040d1ae}
   Action _aGet_Client_exit: Id {bbec42eb-a783-4f5e-82aa-7eeb4cf6f071}
   Action _ainit_active: Id {d9c96ab0-b559-49a2-afe8-ff94a774e454}
   Action _ainit_exit: Id {ad983d6a-a390-4862-a949-8cf9f36606ae}
   Action _ameasure_Deterg_2_active: Id {26827e86-238f-4cae-90ea-080833e3ba15}
   Action _ameasure_Deterg_active: Id {0df3b090-cf38-4d12-bf3b-cbf3c529cdce}
   Action _ameasure_Dis_2_active: Id {1261d4d1-c6d0-4244-bace-be3e25c760cc}
   Action _ameasure_Dis_active: Id {53cb2553-ae2a-4250-8fcc-274b620fda49}
   Action _ameasureDelay_CIP2_1_active: Id {eee92c62-884a-44e9-a331-0195a641ce83}
   Action _ameasureDelay_CIP2_1_entry: Id {5e93bd05-4f42-41e5-8f40-cb8225034977}
   Action _ameasureDelay_CIP2_2_active: Id {e6c27ce5-3263-4596-8180-705d3553666d}
   Action _ameasureDelay_CIP2_2_entry: Id {b1c765b5-bd3e-42f3-a762-17c5119156e5}
   Action _ameasureDelay_CIP4_1_active: Id {95864345-55ce-4583-98e3-3f17b2ed667c}
   Action _ameasureDelay_CIP4_1_entry: Id {f75d6eb0-4cd0-4c37-882c-ed7e1e2ef51d}
   Action _ameasureDelay_CIP4_2_active: Id {79294f20-9c9f-4055-ae02-c5c9b94196a4}
   Action _ameasureDelay_CIP4_2_entry: Id {1aae7665-6957-419b-a173-2f6ea3b229a4}
   Action _aReady_active: Id {560e86d1-cd11-44bd-aed6-a8db9be9b76c}
   Action _aReady_exit: Id {fe06bbde-dba2-4c36-8b83-7a6e8089b6a1}
   Action _aReadyToCondition_Count_active: Id {63783ecf-f88e-4e69-b08a-d0b63a866753}
   Action _aReadyToCondition_Count_entry: Id {c49ce332-1ee4-4760-920c-b0d999acd035}
   Action _aReFill_Water_T93_active: Id {2f420f26-ee2f-4fab-9c41-ff3d506196d6}
   Action _aReFill_Water_T94_active: Id {8d84723c-ae0a-44fc-b26f-f36d0e420f1f}
   Action _aReset_Cond_Tm_CIP2_01_active: Id {93f99ae3-1917-408b-84a5-48debdd15f17}
   Action _aSet_Valves_ToDeafult_active: Id {6f0f9f2b-5faf-4a3e-bc50-2f79008d8530}
   Action _aSet_Valves_ToDeafult_entry: Id {5504b883-dffe-4f34-ad68-2f1bab980d83}
   Action _aSprinkler_Request_CIP1_active: Id {4acc4cf2-f228-4f13-bdcd-db4a92bd7344}
   Action _aSprinkler_Request_CIP35_active: Id {7bbffa29-9878-4026-a507-cc50b1b5b319}
   Action _aStartPump_CIP1_01_active: Id {e50e4f65-8145-4f79-b69c-1a7d9a136df2}
   Action _aStartPump_CIP1_01_entry: Id {d05b04cb-ad28-4d2f-b50e-f58a7739d4a3}
   Action _aStartPump_CIP2_01_active: Id {c1fce140-5edc-4740-a154-cfbe59a57483}
   Action _aStartPump_CIP2_01_entry: Id {4589c8d4-2b8a-47b6-b8e7-d8da9bb4ee5a}
   Action _aStartPump_CIP2_02_active: Id {9ff178c2-f56d-4862-8c8e-bee0c2bafa4c}
   Action _aStartPump_CIP2_02_entry: Id {68002631-498d-4301-be5a-4191a97bd16a}
   Action _aStartPump_CIP2_RPM_01_active: Id {926fdc44-d8f2-4656-9732-79a85aef1568}
   Action _aStartPump_CIP2_RPM_02_active: Id {a603ceb3-2a59-40c6-b08d-10619fb883a4}
   Action _aStartPump_CIP2_RPM_02_entry: Id {e92aaf57-63dd-454d-be83-594290102c87}
   Action _aStartPump_CIP4_RPM_01_active: Id {7055f639-2c8c-427c-8372-ce3721630720}
   Action _aStartPump_CIP4_RPM_02_active: Id {6541b9b3-a926-41a5-a2dd-43356cfd7a84}
   Action _aStartPump_CIP4_01_active: Id {e6aa8b88-0a3e-4980-90b3-b28e3208ca1c}
   Action _aStartPump_CIP4_01_entry: Id {b0df1b3d-bbd7-422e-b23e-87cbef7af745}
   Action _aStartPump_CIP4_02_active: Id {f64d81b7-93d0-4d81-9b19-fca829dbaa54}
   Action _aStartPump_CIP4_02_entry: Id {b59301f9-93ed-4442-a828-b3f5bc9893a8}
   Action _aStartPump_CIP35_active: Id {8f847c4e-380b-4c8e-9efc-5e133107f699}
   Action _aStartPump_CIP35_entry: Id {ce3107e7-d7e1-46a5-b32d-249da89f4251}
   Action _aStop_Pump_entry: Id {48014272-55b2-4c31-adb6-2d01f6affd95}
   Action _aStopPump_CIP1_01_entry: Id {f0260740-b530-49b6-ae60-7945a09e7dde}
   Action _aStopPump_CIP1_02_entry: Id {cf64d467-b785-4967-bf28-6b68d2dc8985}
   Action _aStopPump_CIP2_01_entry: Id {85898c2b-ab66-4edd-b612-16013618240b}
   Action _aStopPump_CIP2_02_entry: Id {df8e1d2d-606f-4c06-afb1-574680199641}
   Action _aStopPump_CIP2_03_entry: Id {0a41a608-f0d9-44c6-a26d-590d4c887acb}
   Action _aStopPump_CIP4_01_entry: Id {f602d6c0-0244-490d-974f-7786e863cb85}
   Action _aStopPump_CIP4_02_entry: Id {6011e812-353e-4927-88db-456a78faf2f5}
   Action _aStopPump_CIP4_03_entry: Id {b282e6dd-a26f-4cdc-82d9-344e825e133b}
   Action _aStopPump_CIP35_01_entry: Id {6a47ecbf-e4c2-4489-963a-6d6de80abe2a}
   Action _aStopPump_CIP35_02_entry: Id {c3d6c7e4-1bec-4f4e-9bfc-b12fa5d63eeb}
   Action _aTank_LowLevel_CIP1_01_active: Id {47975dbe-05c8-4855-a682-02f3a1d90ed0}
   Action _aTank_LowLevel_CIP1_02_active: Id {289829e0-78dc-4147-8ec8-7319f891bc3e}
   Action _aTank_LowLevel_CIP1_02_entry: Id {e7e2eec1-d9c1-47b6-a6d1-cf8acf9c1dc7}
   Action _aTank_LowLevel_CIP2_01_active: Id {58580d6e-e21f-4d3c-a180-0d74f7574119}
   Action _aTank_LowLevel_CIP2_02_active: Id {0b853c55-1b49-4c9f-8a2f-65bb70488411}
   Action _aTank_LowLevel_CIP2_02_entry: Id {a915a083-8ce0-46f9-8f3e-84a27da21374}
   Action _aTank_LowLevel_CIP4_01_active: Id {08010232-500a-48f3-a614-a521a3b4d69c}
   Action _aTank_LowLevel_CIP4_02_active: Id {03ea7d6f-93a1-4a3d-a804-035238dd8a97}
   Action _aTank_LowLevel_CIP4_02_entry: Id {60789d93-6c08-41e6-b874-8551ab513be1}
   Action _aTank_LowLevel_CIP35_01_active: Id {bd1392e8-f7bb-4ffb-a1ec-3aa12b30c399}
   Action _aTank_LowLevel_CIP35_02_active: Id {46b8f49a-c6b6-4094-95d6-c17fbaf2db69}
   Action _aTank_LowLevel_CIP35_02_entry: Id {b05e7121-7b36-4a70-b3fe-4633bbc45de6}
   Action _aTank_MixProof_Clean_CIP2_active: Id {4c83d8fc-5244-4926-8774-0d98cfbda24b}
   Action _aTank_MixProof_Clean_CIP2_entry: Id {3aaabf55-224c-4243-b8e3-e0319731e6c0}
   Action _aTank_MixProof_Clean_CIP4_active: Id {cbf49d17-c130-4e83-9dbe-4bb4a0f1d4a4}
   Action _aTank_MixProof_Clean_CIP4_entry: Id {2430adbb-c9bb-433b-b82a-c79663d4de71}
   Action _aTriBlender_Selection_active: Id {d0e672f4-6afb-4eb1-ae08-259e55e6edbe}
   Action _aTriBlender_Selection_entry: Id {0a68dd9d-1aca-4b6e-aa9d-fe1899267007}
   Action _aWaiting_Client_Drain_Done_active: Id {198d1e9a-548f-4e4c-b425-d71b6a65c8cc}
   Action act_CallProcessControl: Id {ba2500c4-7891-45b7-bd60-804b421a62c3}
   Action act_GetReference: Id {483d260d-ab35-4076-91bc-ffd5a0e6d733}
   Action act_HeatExchng: Id {13b9d6f9-7b3e-4e54-9f53-f81ae43526f9}
   Action act_Oper: Id {c3825564-eb19-4e3f-91a4-377e8a0daffd}
   Action act_ReqBuffer: Id {1b81a7d5-6e97-4216-8c50-f77668c87ac0}
   Action act_Run: Id {1474794e-dde4-4a3c-8164-060b43f4cb22}
   Action act_SprinklerCondition: Id {44149426-1a6f-4c5f-80b5-37350a655a40}
   Method m_Set_CIP_State: Id {f183e936-eac4-4183-abf9-3dd38129926e}
   Method m_DashState_NotAvailable: Id {ef672738-0a06-4f93-93fb-790a43fcc677}
   Method m_Check_ProductionTank_Low_Level: Id {b48f9a03-2e2f-4f01-a8db-812c2687100f}
   Method m_CleanEmpty_Spaces: Id {a02513cf-5921-4270-b511-66d8a68458f2}
   Method m_ClientTank_IsEmpty: Id {b35dd6ac-5e7d-4daa-9425-98b1cad5f40d}
   Method m_ClientTank_Level_IsHigher_Then: Id {8401ba19-06a5-4bdb-9e2e-261fa513b5de}
   Method m_DashState_activate: Id {02085a65-a2cd-4364-8e33-72b46cf78751}
   Method m_DashState_done: Id {7bac3818-529e-4a54-9082-0edd1812249d}
   Method m_DashState_from: Id {517ea0a0-c223-471a-a5e8-76eedc4a5a7a}
   Method m_DashState_Get_ToBeDone_List: Id {d256d03e-5646-4a44-97db-829d1963e250}
   Method m_DashState_Sprinkler: Id {306d9d0f-c147-419d-8576-035700b09af5}
   Method m_DashState_to: Id {90469f15-32d0-4753-bd08-fb0af69e8ea7}
   Method m_DashState_ToString_convertion: Id {ac0b670d-4de4-4707-89c6-0875fdc96ae9}
   Method m_MeasureTimeToHMI: Id {6c49de4b-95a1-4fe1-b1b1-55f4c051916f}
   Method m_OverFlowCorrect: Id {3d927e50-569d-481a-ab49-43c1ca44dff1}
   Method m_PosDelete_HMI: Id {5ecfed30-e439-4aa1-8486-4d270c40480b}
   Method m_PosDeleteAll_HMI: Id {0565b103-e72e-4e42-86f5-de0bd5b6f5d7}
   Method m_PosMove_Down_HMI: Id {c114e84d-a8ed-4e16-9653-147f733c0d8b}
   Method m_PosMove_Up_HMI: Id {882d4194-9591-429b-a6de-feb8c47cbd4c}
   Method m_Set_SFCFlags_Reference: Id {3959a842-c714-4552-9594-b319ee26bb78}
   Method m_TakePosInCIPBuffer: Id {b2dcb157-1d24-4a20-a9df-81a455a5e4d3}
   Method mFillWater: Id {c38e9eb6-e5ec-4b46-a443-d362a1ec1959}
   Method mLoadDefProcessSetPoints: Id {6622ea5b-b543-4ab8-8397-ed9f64ee15e5}
   Method mProcessDeviation: Id {7347b3a8-56cd-4c5d-bbbb-7da59378f31e}
   Method mVolumeMeter: Id {e61a6efb-fd25-4aac-984f-e420c6d353ee}
   Method mVolumeReset_All: Id {90b26673-5b50-4adb-85ab-facca48446ca} *)
